(* IEC 61131-3 sources: PO_LAB_3/Physical/Acp10_MC (part 2) *)

(* ---- acp10_mc.fun ---- *)
FUNCTION_BLOCK MC_AbortTrigger (*aborts FBs connected to trigger events*)
	VAR_INPUT
		Axis : UDINT; (*axis reference, defines on which axis the trigger should be aborted*)
		TriggerInput : MC_TRIGGER_REF; (*trigger input signal source*)
		Execute : BOOL; (*aborts the trigger at rising edge*)
	END_VAR
	VAR_OUTPUT
		Done : BOOL; (*FB with trigger has been aborted*)
		Busy : BOOL; (*the function block is not finished*)
		Error : BOOL; (*error occurred in FB*)
		ErrorID : UINT; (*error number*)
	END_VAR
	VAR
		C_Axis : UDINT; (*internal variable*)
		state : USINT; (*internal variable*)
		C_Done : BOOL; (*internal variable*)
		C_Error : BOOL; (*internal variable*)
		C_ErrorID : UINT; (*internal variable*)
	END_VAR
END_FUNCTION_BLOCK

FUNCTION_BLOCK MC_BR_AutCommand (*transferes commands for the cam automat to the drive*)
	VAR_INPUT
		Slave : UDINT; (*axis reference of the slave axis*)
		Enable : BOOL; (*activates the function block*)
		Start : BOOL; (*starts the cam automat*)
		Stop : BOOL; (*stops the movement on the slave axis*)
		Deceleration : REAL; (*deceleration for the stop command*)
		Restart : BOOL; (*reengages the slave axis to the automat*)
		EndAutomat : BOOL; (*aborts the automat in the background*)
		SetSignal1 : BOOL; (*sets the automat signal1*)
		SetSignal2 : BOOL; (*sets the automat signal2*)
		SetSignal3 : BOOL; (*sets the automat signal3*)
		SetSignal4 : BOOL; (*sets the automat signal4*)
		ResetSignal1 : BOOL; (*resets the automat signal1*)
		ResetSignal2 : BOOL; (*resets the automat signal2*)
		ResetSignal3 : BOOL; (*resets the automat signal3*)
		ResetSignal4 : BOOL; (*resets the automat signal4*)
		TransferParLock : BOOL; (*transfer the par lock parameter*)
		SelectParLock : USINT; (*select the par lock parameter*)
	END_VAR
	VAR_OUTPUT
		Active : BOOL; (*function block is active and waits for command*)
		Busy : BOOL; (*function block is enabled*)
		CommandAborted : BOOL; (*function block was aborted by another function block*)
		Error : BOOL; (*error occurred in the function block*)
		ErrorID : UINT; (*error number*)
		Running : BOOL; (*slave is engaged to the automat*)
		StandBy : BOOL; (*cam automat is active in the background*)
		ParLockTransferred : BOOL; (*par lock parameter transferred*)
		ActualStateIndex : USINT; (*actual state of the cam automat*)
		ActualStateCamIndex : UINT; (*actual cam index of the actual state*)
		InCam : BOOL; (*automat is in cam*)
		InCompensation : BOOL; (*automat is in compensation*)
	END_VAR
	VAR
		C_Slave : UDINT; (*internal variable*)
		IS : MC_0099_IS_TYP; (*internal variable*)
	END_VAR
END_FUNCTION_BLOCK

FUNCTION_BLOCK MC_BR_AutControl (*controls the cam automat functions*)
	VAR_INPUT
		Enable : BOOL; (*enables the functionality of this FB*)
		Slave : UDINT; (*axis reference of the slave axis*)
		ParLock : USINT; (*lock for consistent online change*)
		Signal1 : BOOL; (*set signal1*)
		Signal2 : BOOL; (*set signal2*)
		Signal3 : BOOL; (*set signal3*)
		Signal4 : BOOL; (*set signal4*)
		Start : BOOL; (*start automat*)
		Stop : BOOL; (*stop automat*)
		Deceleration : REAL; (*deceleration for stop command*)
		Restart : BOOL; (*restart command*)
		AdrAutData : UDINT; (*address of optional cam automat data structure*)
		InitAutData : BOOL; (*initialize the parameters of the optional cam automat data structure*)
	END_VAR
	VAR_OUTPUT
		Active : BOOL; (*automat control function block activated*)
		Busy : BOOL; (*function block is not finished*)
		Error : BOOL; (*error occurred in FB*)
		ErrorID : UINT; (*error number*)
		AutDataInitialized : BOOL; (*cam automat data structure initialized*)
		Running : BOOL; (*cam automat is running*)
		ActualStateIndex : USINT; (*index of the actual state*)
		ActualCamType : USINT; (*cam type of the actual state*)
	END_VAR
	VAR
		C_Slave : UDINT; (*internal variable*)
		ParLockOld : USINT; (*internal variable*)
		LockID : USINT; (*internal variable*)
		CmdParLock : BOOL; (*internal variable*)
		EdgeSignal1 : BOOL; (*internal variable*)
		EdgeSignal2 : BOOL; (*internal variable*)
		EdgeSignal3 : BOOL; (*internal variable*)
		EdgeSignal4 : BOOL; (*internal variable*)
		EdgeStart : BOOL; (*internal variable*)
		CmdStart : BOOL; (*internal variable*)
		EdgeStop : BOOL; (*internal variable*)
		CmdStop : BOOL; (*internal variable*)
		C_Deceleration : REAL; (*internal variable*)
		EdgeRestart : BOOL; (*internal variable*)
		CmdRestart : BOOL; (*internal variable*)
		EdgeInitAutData : BOOL; (*internal variable*)
		CmdInitAutData : BOOL; (*internal variable*)
		C_AutData : MC_AUTDATA_TYP; (*internal variable*)
		C_Master : UDINT; (*internal variable*)
		C_Error : BOOL; (*internal variable*)
		C_ErrorID : UINT; (*internal variable*)
		CC_ErrorID : UINT; (*internal variable*)
		SignalSet : USINT; (*internal variable*)
		SignalReset : USINT; (*internal variable*)
		CmdAutStart : UINT; (*internal variable*)
		AutStatusValid : BOOL; (*internal variable*)
		AutStateDld : USINT; (*internal variable*)
		AutStatusOffset : UINT; (*internal variable*)
		AutStatusRecIndex : USINT; (*internal variable*)
		LockIDSend : USINT; (*internal variable*)
		AutActualStateIndexOffset : UINT; (*internal variable*)
		AutActualStateIndexRecIndex : USINT; (*internal variable*)
		C_Busy : BOOL; (*internal variable*)
		AutActualCamTypeOffset : UINT; (*internal variable*)
		AutActualCamTypeRecIndex : USINT; (*internal variable*)
		LockIDMa : USINT; (*internal variable*)
		sendSlot : USINT; (*internal variable*)
		readSlot : USINT; (*internal variable*)
		state : USINT; (*internal variable*)
		LockIDPar : USINT; (*internal variable*)
		MoveID : USINT; (*internal variable*)
		LockIDReceive : USINT; (*internal variable*)
	END_VAR
END_FUNCTION_BLOCK

FUNCTION_BLOCK MC_BR_AutoCamDwell (*starts a link between master and slave with a self calculated cam profile*)
	VAR_INPUT
		Master : UDINT; (*axis reference of the master axis*)
		Slave : UDINT; (*axis reference of the slave axis*)
		Enable : BOOL; (*function block is activated*)
		InitData : BOOL; (*start transferring the parameters*)
		LeadInMasterDistance : REAL; (*master axis compensation distance for the lead in*)
		LeadInSlaveDistance : REAL; (*slave axis compensation distance for the lead in*)
		LeadOutMasterDistance : REAL; (*master axis compensation distance for the lead out*)
		LeadOutSlaveDistance : REAL; (*slave axis compensation distance for the lead out*)
		MasterStartPosition : REAL; (*master position where the cam profile starts*)
		MasterDwellDistance : REAL; (*master length of the optional dwell section*)
		MasterLength : REAL; (*master side length of the automatically calculated cam profile*)
		SlaveLength : REAL; (*slave side length of the automatically calculated cam profile*)
		MasterParID : UINT; (*use this ParID for the master axis instead of the set position*)
		MasterParIDMaxVelocity : REAL; (*maximum speed of the master ParID value*)
		LeadInSignal : BOOL; (*signal from the control to start the lead in*)
		LeadOutSignal : BOOL; (*signal from the control to start the lead out*)
		LeadInParID : UINT; (*ParID that can be used by the drive to start the lead in*)
		LeadOutParID : UINT; (*ParID that can be used by the drive to start the lead out*)
	END_VAR
	VAR_OUTPUT
		Active : BOOL; (*parameters are transferred and FB is active*)
		Busy : BOOL; (*function block is enabled*)
		CommandAborted : BOOL; (*function block aborted by another FB*)
		Error : BOOL; (*error occurred in FB*)
		ErrorID : UINT; (*error number*)
		DataInitialized : BOOL; (*parameters are transferred*)
		InSync : BOOL; (*cam profile is synchronized with the master*)
		InCam : BOOL; (*the coupling is within the cam range*)
		InDwell : BOOL; (*the coupling is within the dwell range*)
	END_VAR
	VAR
		C_Master : UDINT; (*internal variable*)
		C_Slave : UDINT; (*internal variable*)
		EdgeInitData : BOOL; (*internal variable*)
		C_LeadInMasterDistance : DINT; (*internal variable*)
		C_LeadInSlaveDistance : DINT; (*internal variable*)
		C_LeadOutMasterDistance : DINT; (*internal variable*)
		C_LeadOutSlaveDistance : DINT; (*internal variable*)
		C_MasterStartPosition : DINT; (*internal variable*)
		C_MasterDwellDistance : DINT; (*internal variable*)
		C_MasterLength : DINT; (*internal variable*)
		C_SlaveLength : DINT; (*internal variable*)
		C_MasterParID : UINT; (*internal variable*)
		C_MasterParIDMaxVelocity : REAL; (*internal variable*)
		C_LeadInParID : UINT; (*internal variable*)
		C_LeadOutParID : UINT; (*internal variable*)
		EdgeLeadInSignal : BOOL; (*internal variable*)
		EdgeLeadOutSignal : BOOL; (*internal variable*)
		LeadInSignalUsed : BOOL; (*internal variable*)
		LeadOutSignalUsed : BOOL; (*internal variable*)
		C_Active : BOOL; (*internal variable*)
		C_Busy : BOOL; (*internal variable*)
		C_CommandAborted : BOOL; (*internal variable*)
		C_Error : BOOL; (*internal variable*)
		C_ErrorID : UINT; (*internal variable*)
		CC_ErrorID : UINT; (*internal variable*)
		C_InSync : BOOL; (*internal variable*)
		C_InCam : BOOL; (*internal variable*)
		C_InDwell : BOOL; (*internal variable*)
		RunningMasterDwellDistance : DINT; (*internal variable*)
		ArithIndex : UINT; (*internal variable*)
		CmpIndex : UINT; (*internal variable*)
		MuxIndex : UINT; (*internal variable*)
		EvWrIndex : UINT; (*internal variable*)
		VarIndex : UINT; (*internal variable*)
		LogicIndex : UINT; (*internal variable*)
		AutStatusValid : BOOL; (*internal variable*)
		AutActualStateIndexOffset : UINT; (*internal variable*)
		AutActualStateIndexRecIndex : USINT; (*internal variable*)
		LockIDMa : USINT; (*internal variable*)
		sendSlot : USINT; (*internal variable*)
		readSlot : USINT; (*internal variable*)
		state : USINT; (*internal variable*)
		LockID : USINT; (*internal variable*)
		LockIDPar : USINT; (*internal variable*)
		LockIDSend : USINT; (*internal variable*)
		MoveID : USINT; (*internal variable*)
		LockIDReceive : USINT; (*internal variable*)
	END_VAR
END_FUNCTION_BLOCK

FUNCTION_BLOCK MC_BR_AxisErrorCollector (*collects information if a FB or axis error occured and if an axis is in state Errorstop*)
	VAR_INPUT
		Axis : UDINT; (*axis reference*)
		Enable : BOOL; (*function block is activated*)
	END_VAR
	VAR_OUTPUT
		Valid : BOOL; (*if set, the data of the other outputs is valid*)
		Busy : BOOL; (*function block is not finished*)
		Error : BOOL; (*error occurred in FB*)
		ErrorID : UINT; (*error number*)
		FunctionBlockError : BOOL; (*at least one function block reported an error*)
		AxisError : BOOL; (*at least one axis error was reported*)
		AxisWarning : BOOL; (*at least one axis warning was reported*)
		Errorstop : BOOL; (*the axis is in state Errorstop*)
	END_VAR
	VAR
		C_Axis : UDINT; (*internal variable*)
		IS : MC_0104_IS_TYP; (*internal variable*)
	END_VAR
END_FUNCTION_BLOCK

FUNCTION_BLOCK MC_BR_BrakeControl (*executes several commands for holding brake*)
	VAR_INPUT
		Axis : UDINT; (*axis reference*)
		Execute : BOOL; (*execute brake command at rising edge*)
		Command : USINT; (*brake command*)
		Configuration : MC_BRAKE_CONFIG_REF; (*brake configuration*)
	END_VAR
	VAR_OUTPUT
		Done : BOOL; (*brake command done*)
		Busy : BOOL; (*function block is not finished*)
		Error : BOOL; (*error occured in FB*)
		ErrorID : UINT; (*error number*)
		PositionError : REAL; (*position error of holding brake test*)
		BrakeStatus : BOOL; (*actual brake status*)
	END_VAR
	VAR
		C_Axis : UDINT; (*internal variable*)
		IS : MC_0110_IS_TYP; (*internal variable*)
	END_VAR
END_FUNCTION_BLOCK

FUNCTION_BLOCK MC_BR_BrakeOperation (*opens and closes the holding brake when the controller is off*)
	VAR_INPUT
		Axis : UDINT; (*axis reference*)
		Execute : BOOL; (*execute brake command at rising edge*)
		BrakeCommand : USINT; (*brake command, open or close*)
	END_VAR
	VAR_OUTPUT
		Done : BOOL; (*brake command done*)
		Busy : BOOL; (*function block is not finished*)
		Error : BOOL; (*error occurred in FB*)
		ErrorID : UINT; (*error number*)
	END_VAR
	VAR
		C_Axis : UDINT; (*internal variable*)
		C_Execute : BOOL; (*internal variable*)
		C_BrakeCommand : USINT; (*internal variable*)
		C_Done : BOOL; (*internal variable*)
		LockIDPar : USINT; (*internal variable*)
		C_ErrorID : UINT; (*internal variable*)
		C_Error : BOOL; (*internal variable*)
		state : USINT; (*internal variable*)
	END_VAR
END_FUNCTION_BLOCK

FUNCTION_BLOCK MC_BR_CalcCamFromPoints (*calculates a cam profile from a list of points*)
	VAR_INPUT
		Execute : BOOL; (*calculation starts at rising edge*)
		MasterPointsAddress : UDINT; (*data address of the master points list*)
		SlavePointsAddress : UDINT; (*data address of the slave points list*)
		NumberOfPoints : UINT; (*number of master and slave points*)
		CamProfileAddress : UDINT; (*data address for the calculated cam profile*)
		Configuration : MC_CALC_CAM_CONFIG_REF; (*optional additional configuration*)
	END_VAR
	VAR_OUTPUT
		Done : BOOL; (*calculation is complete*)
		Busy : BOOL; (*function block is not finished*)
		Error : BOOL; (*error occurred in FB*)
		ErrorID : UINT; (*error number*)
	END_VAR
	VAR
		IS : MC_0093_IS_TYP; (*internal variable*)
	END_VAR
END_FUNCTION_BLOCK

FUNCTION_BLOCK MC_BR_CalcCamFromSections (*calculates from a list of points a cam profile*)
	VAR_INPUT
		Execute : BOOL; (*calculation starts at rising edge*)
		DataAddress : UDINT; (*data address of the input data with the list of points*)
		CamProfileAddress : UDINT; (*data address for the calculated cam profile*)
	END_VAR
	VAR_OUTPUT
		Done : BOOL; (*calculation is complete*)
		Busy : BOOL; (*function block is not finished*)
		Error : BOOL; (*error occurred in FB*)
		ErrorID : UINT; (*error number*)
		ErrorInSection : UINT; (*index of section with error*)
	END_VAR
	VAR
		C_ErrorID : UINT; (*internal variable*)
		C_ErrorInSection : UINT; (*internal variable*)
		C_Error : BOOL; (*internal variable*)
		state : USINT; (*internal variable*)
	END_VAR
END_FUNCTION_BLOCK

FUNCTION_BLOCK MC_BR_CalcPointsFromCam (*calculates a list of points from a cam profile*)
	VAR_INPUT
		Execute : BOOL; (*calculation starts at rising edge*)
		DataObjectName : STRING[12]; (*name of the cam table*)
		MasterPointsAddress : UDINT; (*data address of the master points list*)
		SlavePointsAddress : UDINT; (*data address of the slave points list*)
		NumberOfPoints : UINT; (*number of master and slave points*)
	END_VAR
	VAR_OUTPUT
		Done : BOOL; (*calculation is complete*)
		Busy : BOOL; (*function block is not finished *)
		Error : BOOL; (*error occured in FB*)
		ErrorID : UINT; (*error number*)
		AdditionalInfo : MC_CALC_CAM_CONFIG_REF; (*additional information about the cam profile*)
	END_VAR
	VAR
		IS : MC_0123_IS_TYP; (*internal variable*)
	END_VAR
END_FUNCTION_BLOCK

FUNCTION_BLOCK MC_BR_CalcSectionsFromCam (*calculates the sections from a cam profile *)
	VAR_INPUT
		Execute : BOOL; (*calculation starts at rising edge*)
		DataObjectName : STRING[12]; (*name of the cam table*)
		DataAddress : UDINT; (*address of the variable for the sections*)
	END_VAR
	VAR_OUTPUT
		Done : BOOL; (*calculation is complete*)
		Busy : BOOL; (*function block is not finished *)
		Error : BOOL; (*error occured in FB*)
		ErrorID : UINT; (*error number*)
	END_VAR
	VAR
		IS : MC_0122_IS_TYP; (*internal variable*)
	END_VAR
END_FUNCTION_BLOCK

FUNCTION_BLOCK MC_BR_CamIn (*starts a cam profile link between the master and the slave axis*)
	VAR_INPUT
		Master : UDINT; (*axis reference of the master axis*)
		Slave : UDINT; (*axis reference of the slave axis*)
		Enable : BOOL; (*function block is activated*)
		InitData : BOOL; (*starts transferring the parameters*)
		CamTableID : USINT; (*ID number of the cam profile*)
		MasterStartPosition : REAL; (*master position where the cam profile starts*)
		MasterScaling : DINT; (*factor of the master profile*)
		SlaveScaling : DINT; (*factor of the slave scaling*)
		EnterCam : BOOL; (*signal from the control to start the coupling*)
		ExitCam : BOOL; (*signal from the control to end the coupling*)
		Restart : BOOL; (*signal from the control to restart the coupling*)
        AdvancedParameters: MC_ADVANCED_CAM_PAR_REF; (*additional inputs for advanced usage of FB*)
	END_VAR
	VAR_OUTPUT
		Active : BOOL; (*parameters are transferred and FB is active*)
		Busy : BOOL; (*function block is enabled*)
		CommandAborted : BOOL; (*function block aborted by another FB*)
		Error : BOOL; (*error occurred in FB*)
		ErrorID : UINT; (*error number*)
		DataInitialized : BOOL; (*transferring parameters is completed*)
		Running : BOOL; (*cam coupling is running*)
		StandBy : BOOL; (*cam coupling is active in the background*)
		InLeadIn : BOOL; (*the coupling is within the leadin range*)
		InCam : BOOL; (*the coupling is within the cam range*)
		InLeadOut : BOOL; (*the coupling is within the leadout range*)
		EndOfProfile : BOOL; (*pulsed output signaling the cyclic end of the cam profile*)
	END_VAR
	VAR
		C_Master : UDINT; (*internal variable*)
		C_Slave : UDINT; (*internal variable*)
		IS: MC_0146_IS_TYP; (*internal variable*)
	END_VAR
END_FUNCTION_BLOCK

FUNCTION_BLOCK MC_BR_CamDwell (*starts a cam profile link between the master and the slave axis*)
	VAR_INPUT
		Master : UDINT; (*axis reference of the master axis*)
		Slave : UDINT; (*axis reference of the slave axis*)
		Enable : BOOL; (*function block is activated*)
		InitData : BOOL; (*starts transferring the parameters*)
		LeadInMasterDistance : REAL; (*master axis compensation distance for the lead in*)
		LeadInSlaveDistance : REAL; (*slave axis compensation distance for the lead in*)
		LeadInMasterOffset : REAL; (*master side offset within the cam profile*)
		LeadOutMasterDistance : REAL; (*master axis compensation distance for the lead out*)
		LeadOutSlaveDistance : REAL; (*slave axis compensation distance for the lead out*)
		LeadOutMasterOffset : REAL; (*master side offset within the cam profile*)
		MasterStartPosition : REAL; (*master position where the cam profile starts*)
		MasterDwellDistance : REAL; (*master length of the optional dwell section*)
		MasterScaling : REAL; (*factor of the master profile*)
		SlaveScaling : REAL; (*factor of the slave scaling*)
		CamTableID : USINT; (*ID number of the cam profile*)
		MasterParID : UINT; (*use this ParID for the master axis instead of the set position*)
		MasterParIDMaxVelocity : REAL; (*maximum speed of the master ParID value*)
		LeadInSignal : BOOL; (*signal from the control to start the lead in*)
		LeadOutSignal : BOOL; (*signal from the control to start the lead out*)
		LeadInParID : UINT; (*ParID that can be used by the drive to start the lead out movement*)
		LeadOutParID : UINT; (*ParID that can be used by the drive to start the lead out movement*)
	END_VAR
	VAR_OUTPUT
		Active : BOOL; (*parameters are transferred and FB is active*)
		Busy : BOOL; (*function block is enabled*)
		CommandAborted : BOOL; (*function block aborted by another FB*)
		Error : BOOL; (*error occurred in FB*)
		ErrorID : UINT; (*error number*)
		DataInitialized : BOOL; (*transferring parameters is completed*)
		InSync : BOOL; (*cam profile is synchronized with the master*)
		InCam : BOOL; (*the coupling is within the cam range*)
		InDwell : BOOL; (*the coupling is within the dwell range*)
	END_VAR
	VAR
		C_Master : UDINT; (*internal variable*)
		C_Slave : UDINT; (*internal variable*)
		EdgeInitData : BOOL; (*internal variable*)
		C_LeadInMasterDistance : DINT; (*internal variable*)
		C_LeadInSlaveDistance : DINT; (*internal variable*)
		C_LeadInMasterOffset : DINT; (*internal variable*)
		C_LeadOutMasterDistance : DINT; (*internal variable*)
		C_LeadOutSlaveDistance : DINT; (*internal variable*)
		C_LeadOutMasterOffset : DINT; (*internal variable*)
		C_MasterStartPosition : DINT; (*internal variable*)
		C_MasterDwellDistance : DINT; (*internal variable*)
		C_MasterScaling : DINT; (*internal variable*)
		C_SlaveScaling : DINT; (*internal variable*)
		C_CamTableID : UINT; (*internal variable*)
		C_MasterParID : UINT; (*internal variable*)
		C_MasterParIDMaxVelocity : REAL; (*internal variable*)
		C_LeadInParID : UINT; (*internal variable*)
		C_LeadOutParID : UINT; (*internal variable*)
		EdgeLeadInSignal : BOOL; (*internal variable*)
		EdgeLeadOutSignal : BOOL; (*internal variable*)
		LeadInSignalUsed : BOOL; (*internal variable*)
		LeadOutSignalUsed : BOOL; (*internal variable*)
		C_Active : BOOL; (*internal variable*)
		C_Busy : BOOL; (*internal variable*)
		C_CommandAborted : BOOL; (*internal variable*)
		C_Error : BOOL; (*internal variable*)
		C_ErrorID : UINT; (*internal variable*)
		CC_ErrorID : UINT; (*internal variable*)
		C_InSync : BOOL; (*internal variable*)
		C_InCam : BOOL; (*internal variable*)
		C_InDwell : BOOL; (*internal variable*)
		RunningMasterDwellDistance : DINT; (*internal variable*)
		ArithIndex : UINT; (*internal variable*)
		CmpIndex : UINT; (*internal variable*)
		MuxIndex : UINT; (*internal variable*)
		EvWrIndex : UINT; (*internal variable*)
		VarIndex : UINT; (*internal variable*)
		LogicIndex : UINT; (*internal variable*)
		AutStatusValid : BOOL; (*internal variable*)
		AutActualStateIndexOffset : UINT; (*internal variable*)
		AutActualStateIndexRecIndex : USINT; (*internal variable*)
		LockIDMa : USINT; (*internal variable*)
		AutActualCamTypeOffset : UINT; (*internal variable*)
		AutActualCamTypeRecIndex : USINT; (*internal variable*)
		LockIDSend : USINT; (*internal variable*)
		sendSlot : USINT; (*internal variable*)
		readSlot : USINT; (*internal variable*)
		state : USINT; (*internal variable*)
		LockID : USINT; (*internal variable*)
		LockIDPar : USINT; (*internal variable*)
		LockIDReceive : USINT; (*internal variable*)
		MoveID : USINT; (*internal variable*)
	END_VAR
END_FUNCTION_BLOCK

FUNCTION_BLOCK MC_BR_CamTransition (*starts a cam profile link between the master and the slave axis*)
	VAR_INPUT
		Master : UDINT; (*axis reference of the master axis*)
		Slave : UDINT; (*axis reference of the slave axis*)
		Enable : BOOL; (*function block is activated*)
		InitData : BOOL; (*starts transferring the parameters*)
		LeadInMasterDistance : REAL; (*master axis compensation distance for the lead in*)
		LeadInSlaveDistance : REAL; (*slave axis compensation distance for the lead in*)
		LeadInMasterOffset : REAL; (*master side offset within the cam profile*)
		LeadOutMasterDistance : REAL; (*master axis compensation distance for the lead out*)
		LeadOutSlaveDistance : REAL; (*slave axis compensation distance for the lead out*)
		LeadOutMasterOffset : REAL; (*master side offset within the cam profile*)
		ReverseSlaveDistance : REAL; (*slaves moves this distence in reverse direction during transition*)
		MasterInterval : REAL; (*interval length of master movement: cam + transition*)
		SlaveInterval : REAL; (*interval length of slave movement: cam + transition*)
		MasterStartPosition : REAL; (*master position where the cam profile starts*)
		MasterScaling : REAL; (*factor of the master profile*)
		SlaveScaling : REAL; (*factor of the slave scaling*)
		CamTableID : USINT; (*ID number of the cam profile*)
		MasterParID : UINT; (*use this ParID for the master axis instead of the set position*)
		MasterParIDMaxVelocity : REAL; (*maximum speed of the master ParID value*)
		LeadInSignal : BOOL; (*signal from the control to start the lead in*)
		LeadOutSignal : BOOL; (*signal from the control to start the lead out*)
		LeadInParID : UINT; (*ParID that can be used by the drive to start the lead out movement*)
		LeadOutParID : UINT; (*ParID that can be used by the drive to start the lead out movement*)
		TransitionMode : UINT; (*mode for transition movement*)
		CamMode : UINT; (*mode for cam movement*)
		CamTime : REAL; (*time for cam movement in mode mcTIME_BASED*)
	END_VAR
	VAR_OUTPUT
		Active : BOOL; (*parameters are transferred and FB is active*)
		Busy : BOOL; (*function block is enabled*)
		CommandAborted : BOOL; (*function block aborted by another FB*)
		Error : BOOL; (*error occurred in FB*)
		ErrorID : UINT; (*error number*)
		DataInitialized : BOOL; (*transferring parameters is completed*)
		InSync : BOOL; (*cam profile is synchronized with the master*)
		InLeadIn : BOOL; (*the coupling is within the leadin range*)
		InCam : BOOL; (*the coupling is within the cam range*)
		InTransition : BOOL; (*the coupling is within the transition range*)
		InReverse : BOOL; (*the coupling is within the reverse reange*)
		InLeadOut : BOOL; (*the coupling is within the leadout range*)
	END_VAR
	VAR
		C_Master : UDINT; (*internal variable*)
		C_Slave : UDINT; (*internal variable*)
		EdgeInitData : BOOL; (*internal variable*)
		C_LeadInMasterDistance : DINT; (*internal variable*)
		C_LeadInSlaveDistance : DINT; (*internal variable*)
		C_LeadInMasterOffset : DINT; (*internal variable*)
		C_LeadOutMasterDistance : DINT; (*internal variable*)
		C_LeadOutSlaveDistance : DINT; (*internal variable*)
		C_LeadOutMasterOffset : DINT; (*internal variable*)
		C_ReverseSlaveDistance : DINT; (*internal variable*)
		C_MasterInterval : DINT; (*internal variable*)
		C_SlaveInterval : DINT; (*internal variable*)
		C_MasterStartPosition : DINT; (*internal variable*)
		C_MasterScaling : DINT; (*internal variable*)
		C_SlaveScaling : DINT; (*internal variable*)
		C_CamTableID : UINT; (*internal variable*)
		C_MasterParID : UINT; (*internal variable*)
		C_MasterParIDMaxVelocity : REAL; (*internal variable*)
		C_LeadInParID : UINT; (*internal variable*)
		C_LeadOutParID : UINT; (*internal variable*)
		C_TransitionMode : UINT; (*internal variable*)
		C_CamMode : UINT; (*internal variable*)
		C_CamTime : REAL; (*internal variable*)
		EdgeLeadInSignal : BOOL; (*internal variable*)
		EdgeLeadOutSignal : BOOL; (*internal variable*)
		LeadInSignalUsed : BOOL; (*internal variable*)
		LeadOutSignalUsed : BOOL; (*internal variable*)
		C_Active : BOOL; (*internal variable*)
		C_Busy : BOOL; (*internal variable*)
		C_CommandAborted : BOOL; (*internal variable*)
		C_Error : BOOL; (*internal variable*)
		C_ErrorID : UINT; (*internal variable*)
		CC_ErrorID : UINT; (*internal variable*)
		C_InSync : BOOL; (*internal variable*)
		C_InCam : BOOL; (*internal variable*)
		C_InTransition : BOOL; (*internal variable*)
		C_InReverse : BOOL; (*internal variable*)
		C_InLeadIn : BOOL; (*internal variable*)
		C_InLeadOut : BOOL; (*internal variable*)
		C_MasterCompDistance : DINT; (*internal variable*)
		C_SlaveCompDistance : DINT; (*internal variable*)
		C_OldMasterCompDistance : DINT; (*internal variable*)
		C_OldSlaveCompDistance : DINT; (*internal variable*)
		C_CamMasterPeriod : DINT; (*internal variable*)
		C_CamSlavePeriod : DINT; (*internal variable*)
		ArithIndex : UINT; (*internal variable*)
		CmpIndex : UINT; (*internal variable*)
		MuxIndex : UINT; (*internal variable*)
		EvWrIndex : UINT; (*internal variable*)
		VarIndex : UINT; (*internal variable*)
		LogicIndex : UINT; (*internal variable*)
		PidIndex : UINT; (*internal variable*)
		AutStatusValid : BOOL; (*internal variable*)
		InitDataUsed : BOOL; (*internal variable*)
		AutActualStateIndexOffset : UINT; (*internal variable*)
		AutActualStateIndexRecIndex : USINT; (*internal variable*)
		oldAutomatState : USINT; (*internal variable*)
		MasterVelocityOffset : UINT; (*internal variable*)
		MasterVelocityRecIndex : USINT; (*internal variable*)
		LockIDMa : USINT; (*internal variable*)
		AutActualCamTypeOffset : UINT; (*internal variable*)
		AutActualCamTypeRecIndex : USINT; (*internal variable*)
		ChangePending : BOOL; (*internal variable*)
		sendSlot : USINT; (*internal variable*)
		readSlot : USINT; (*internal variable*)
		state : USINT; (*internal variable*)
		LockID : USINT; (*internal variable*)
		LockIDPar : USINT; (*internal variable*)
		MoveID : USINT; (*internal variable*)
		LockIDSend : USINT; (*internal variable*)
		Reserve3 : UDINT; (*internal variable*)
		nextState : USINT; (*internal variable*)
		Reserve4 : USINT; (*internal variable*)
		LockIDReceive : USINT; (*internal variable*)
		Reserve6 : BOOL; (*internal variable*)
	END_VAR
END_FUNCTION_BLOCK

FUNCTION_BLOCK MC_BR_CheckAutCompensation (*checks the compensation data of a cam profile automat*)
	VAR_INPUT
		Master : UDINT; (*axis reference of the master axis*)
		Slave : UDINT; (*axis reference of the slave axis*)
		Execute : BOOL; (*check the compensation data at rising edge*)
		Mode : UINT; (*choose the mode*)
		CompensationData : MC_AUT_COMP_DATA_REF; (*compensation data for the check or calculation*)
	END_VAR
	VAR_OUTPUT
		Done : BOOL; (*check or calculation is successfully finished*)
		Busy : BOOL; (*function block is not finished yet*)
		Error : BOOL; (*error occured in FB*)
		ErrorID : UINT; (*error number*)
		Result : REAL; (*result of the calculation*)
	END_VAR
	VAR
		C_Master : UDINT; (*internal variable*)
		C_Slave : UDINT; (*internal variable*)
		IS : MC_0103_IS_TYP; (*internal variable*)
	END_VAR
END_FUNCTION_BLOCK

FUNCTION_BLOCK MC_BR_CheckEndlessPosition (*checks the endless position data for restoring the axis position*)
	VAR_INPUT
		Axis : UDINT; (*axis reference*)
		Execute : BOOL; (*check the endless position data at rising edge*)
		DataAddress : UDINT; (*data address of momory storage for endless position*)
	END_VAR
	VAR_OUTPUT
		Done : BOOL; (*memory storage for endless position was checked*)
		Busy : BOOL; (*function block is not finished*)
		Error : BOOL; (*error occurred in FB*)
		ErrorID : UINT; (*error number*)
		EndlessPositionInitialized : BOOL; (*address of memory storage already initialized*)
		DataValid : BOOL; (*axis position can be restored from the endless position data*)
	END_VAR
	VAR
		C_Axis : UDINT; (*internal variable*)
		IS : MC_0130_IS_TYP; (*internal variable*)
	END_VAR
END_FUNCTION_BLOCK

FUNCTION_BLOCK MC_BR_CommandError (*transfers error commands to the drive, where they are entered*)
	VAR_INPUT
		Axis  : UDINT; (*axis reference*)
		Execute : BOOL; (*transfer command at rising edge*)
		Command : UINT; (*error command*)
	END_VAR
	VAR_OUTPUT
		Done  : BOOL; (*command was successfully transferred *)
		Busy  : BOOL; (*function block is not finished yet*)
		Error : BOOL; (*error occured in FB*)
		ErrorID : UINT; (*error number *)
	END_VAR
	VAR
		C_Axis : UDINT; (*internal variable*)
		IS : MC_0140_IS_TYP; (*internal variable*)
	END_VAR
END_FUNCTION_BLOCK

FUNCTION_BLOCK MC_BR_ConfigPowerStageCheck (*configurates the power stage checks of the ACOPOS*)
	VAR_INPUT
		Axis : UDINT; (*axis reference*)
		Execute : BOOL; (*transfer configuration at rising edge *)
		Configuration : MC_POWER_STAGE_CHECK_REF; (*configuration data*)
	END_VAR
	VAR_OUTPUT
		Done : BOOL; (*configuration is successfully finished*)
		Busy : BOOL; (*function block is not finished yet*)
		Error : BOOL; (*error occured in FB*)
		ErrorID : UINT; (*error number*)
	END_VAR
	VAR
		C_Axis : UDINT; (*internal variable*)
		IS : MC_0137_IS_TYP; (*internal variable*)
	END_VAR
END_FUNCTION_BLOCK

FUNCTION_BLOCK MC_BR_CrossCutterControl (*controls a cutter axis linked to a master axis*)
	VAR_INPUT
		Master : UDINT; (*axis reference of the master axis*)
		Slave : UDINT; (*axis reference of the slave/cutter axis*)
		Enable : BOOL; (*function block is activated*)
		InitData : BOOL; (*starts transferring the parameters*)
		EnableCut : BOOL; (*start/stop synchronizing slave to master*)
		CutRangeMaster : REAL; (*cut area on master axis, where the cutter needs to run synchronous to master*)
		CutRangeSlave : REAL; (*area around cut point on slave axis, where the cutter needs to run synchronous to master*)
		ProductLength : REAL; (*distance (master based) in which the cutter needs to make one cut*)
		ProductLengthCorrection : REAL; (*this value is added to ProductLength and then downloaded*)
		AdvancedParameters : MC_ADVANCED_CUT_PAR_REF; (*additional inputs for advanced usage of FB*)
	END_VAR
	VAR_OUTPUT
		Active : BOOL; (*parameters are transferred and FB is active*)
		Busy : BOOL; (*function block is enabled*)
		CommandAborted : BOOL; (*function block aborted by another FB*)
		Error : BOOL; (*error occurred in FB*)
		ErrorID : UINT; (*error number*)
		DataInitialized : BOOL; (*transferring parameters is completed*)
		StandBy : BOOL; (*FB can be restarted*)
		InCompensation : BOOL; (*axis outside CutRange, and synchronized*)
		InCut : BOOL; (*axis is within CutRange*)
		CutCount : UDINT; (*information about how many cuts have been made*)
		CutMasterPosition : DINT; (*latched master position at cut for registration mark control*)
	END_VAR
	VAR
		C_Master : UDINT; (*internal variable*)
		C_Slave : UDINT; (*internal variable*)
		IS : MC_0114_IS_TYP; (*internal variable*)
	END_VAR
END_FUNCTION_BLOCK

FUNCTION_BLOCK MC_BR_CyclicRead (*enters the specified ParID in the cyclic data from drive and returns it*)
	VAR_INPUT
		Axis : UDINT; (*axis reference*)
		Enable : BOOL; (*specified ParID is read from the drive as long as enable is TRUE*)
		ParID : UINT; (*ParID which should be read from the drive*)
		DataAddress : UDINT; (*data address of the variable for the value of the ParID*)
		DataType : UINT; (*data type of the ParID*)
		Mode : UINT; (*mode for configuration of records*)
	END_VAR
	VAR_OUTPUT
		Valid : BOOL; (*when set the output is valid*)
		Busy : BOOL; (*function block is not finished*)
		Error : BOOL; (*error occurred in FB*)
		ErrorID : UINT; (*error number*)
	END_VAR
	VAR
		C_Axis : UDINT; (*internal variable*)
		IS : MC_0069_IS_TYP; (*internal variable*)
	END_VAR
END_FUNCTION_BLOCK

FUNCTION_BLOCK MC_BR_CyclicReadDataInfo (*Read administrative information of cyclic read data*)
	VAR_INPUT
		Axis : UDINT; (*axis reference*)
		Enable : BOOL; (*function block is activated*)
	END_VAR
	VAR_OUTPUT
		Valid : BOOL; (*if set, the data of the other outputs is valid*)
		Busy : BOOL; (*function block is not finished*)
		Error : BOOL; (*error occurred in FB*)
		ErrorID : UINT; (*error number*)
		RecordCount : UINT; (*number of configured records from the drive*)
		ParIDCount : UINT; (*number of configured ParIDs from the drive*)
		RecordUpdateTime : DINT; (*update time of one single record from the drive*)
		TotalUpdateTime : DINT; (*update time of all records from the drive*)
		RecordIndex : UINT; (*index of currently read record from the drive*)
		RecordInfo : MC_RECORD_INFO_REF; (*detailed information about all records from the drive*)
	END_VAR
	VAR
		C_Axis : UDINT; (*internal variable*)
		IS : MC_0098_IS_TYP; (*internal structure*)
	END_VAR
END_FUNCTION_BLOCK

FUNCTION_BLOCK MC_BR_CyclicWrite (*enters a specified ParID in the cyclic data to drive*)
	VAR_INPUT
		Axis : UDINT; (*axis reference*)
		Enable : BOOL; (*specified ParID is written to the drive as long as enable is TRUE*)
		ParID : UINT; (*ParID which should be written to the drive*)
		DataAddress : UDINT; (*data address of the variable with the value for the ParID*)
		DataType : UINT; (*data type of the ParID*)
		Mode : UINT; (*currently not used*)
	END_VAR
	VAR_OUTPUT
		Valid : BOOL; (*when set the output is valid*)
		Busy : BOOL; (*function block is not finished*)
		Error : BOOL; (*error occurred in FB*)
		ErrorID : UINT; (*error number*)
	END_VAR
	VAR
		C_Axis : UDINT; (*internal variable*)
		IS : MC_0070_IS_TYP; (*internal variable*)
	END_VAR
END_FUNCTION_BLOCK

FUNCTION_BLOCK MC_BR_DigitalCamSwitch (*allows a digital output (Track) to be set whenever the axis is inside a position window*)
	VAR_INPUT
		Enable : BOOL; (*when set the FB parameters are downloaded*)
		Switches : MC_MASTER_SWITCHES_REF; (*reference to the switching actions*)
		OutputOptions : MC_OUTPUT_OPTIONS_REF; (*reference to the output options*)
		TrackOptions : MC_TRACK_OPTIONS_REF; (*reference to the track options*)
		SwitchSelector : USINT; (*selection of the switching data*)
		EnableValue : BOOL; (*enable the output of the state of the track on the FB output*)
		EnableParID : BOOL; (*enable the output of the state of the track on the specified ParID*)
		EnableDigOut : BOOL; (*enable the output of of the state of the track on a plug-in module*)
		ChangeSwitches : BOOL; (*change the active switching data*)
		InitSwitches : BOOL; (*initialize new switching parameters*)
		InitTrackOptions : BOOL; (*initialize new track options*)
	END_VAR
	VAR_OUTPUT
		InOperation : BOOL; (*is set after all parameters are transferred*)
		Busy : BOOL; (*the function block is active*)
		Error : BOOL; (*error occured in FB*)
		ErrorID : UINT; (*error number*)
		SwitchesChanged : BOOL; (*the active switching data has been changed*)
		SwitchesInitialized : BOOL; (*new switching parameters are initialized*)
		TrackOptionsInitialized : BOOL; (*new track options initialized*)
		Value : BOOL; (*actual state of the track*)
		ActualSwitches : USINT; (*actual active switches*)
	END_VAR
	VAR
		IS : MC_0107_IS_TYP; (*internal variable*)
		C_Master : UDINT; (*internal variable*)
		C_Slave : UDINT; (*internal variable*)
	END_VAR
END_FUNCTION_BLOCK

FUNCTION_BLOCK MC_BR_DownloadCamProfileObj (*transfers a cam profile object to the drive*)
	VAR_INPUT
		Axis : UDINT; (*axis reference*)
		Execute : BOOL; (*download camprofile at rising edge*)
		DataObjectName : STRING[12]; (*name of the data object*)
		Index : UINT; (*index for cam profile data object*)
		Periodic : BOOL; (*select if paeriodic or non periodic*)
	END_VAR
	VAR_OUTPUT
		Done : BOOL; (*download completed*)
		Busy : BOOL; (*function block is not finished*)
		Error : BOOL; (*error occurred in FB*)
		ErrorID : UINT; (*error number*)
	END_VAR
	VAR
		C_Axis : UDINT; (*internal variable*)
		C_DataObjectName : STRING[12]; (*internal variable*)
		LockIDPar : USINT; (*internal variable*)
		C_Error : BOOL; (*internal variable*)
		C_Index : UINT; (*internal variable*)
		C_ErrorID : UINT; (*internal variable*)
		C_Periodic : BOOL; (*internal variable*)
		C_Done : BOOL; (*internal variable*)
		state : USINT; (*internal variable*)
	END_VAR
END_FUNCTION_BLOCK

FUNCTION_BLOCK MC_BR_DownloadCamProfileData (*transfers cam profile data to the drive*)
	VAR_INPUT
		Axis : UDINT; (*axis reference*)
		Execute : BOOL; (*download cam profile at rising edge*)
		DataAddress : UDINT; (*address of cam profile data*)
		Index : UINT; (*index for cam profile data object*)
		Periodic : BOOL; (*decides if periodic or not*)
	END_VAR
	VAR_OUTPUT
		Done : BOOL; (*download completed*)
		Busy : BOOL; (*function block is not fnished*)
		Error : BOOL; (*error occurred in FB*)
		ErrorID : UINT; (*error number*)
	END_VAR
	VAR
		C_Axis : UDINT; (*internal variable*)
		C_DataAddress : UDINT; (*internal variable*)
		C_Index : UINT; (*internal variable*)
		C_ErrorID : UINT; (*internal variable*)
		C_Error : BOOL; (*internal variable*)
		C_Periodic : BOOL; (*internal variable*)
		C_Done : BOOL; (*internal variable*)
		state : USINT; (*internal variable*)
		LockIDPar : USINT; (*internal variable*)
	END_VAR
END_FUNCTION_BLOCK

FUNCTION_BLOCK MC_BR_DownloadParSequ (*downloads a parameter sequence*)
	VAR_INPUT
		Axis : UDINT; (*axis reference*)
		Execute : BOOL; (*download parameter sequence at rising edge*)
		DataAddress : UDINT; (*data address of the parameter sequence*)
	END_VAR
	VAR_OUTPUT
		Done : BOOL; (*download completed*)
		Busy : BOOL; (*function block is not finished*)
		Error : BOOL; (*error occurred*)
		ErrorID : UINT; (*error number*)
	END_VAR
	VAR
		Reserve1 : UINT; (*internal variable*)
		C_Axis : UDINT; (*internal variable*)
		C_DataAddress : UDINT; (*internal variable*)
		C_Done : BOOL; (*internal variable*)
		C_Error : BOOL; (*internal variable*)
		C_ErrorID : UINT; (*internal variable*)
		LockIDPar : USINT; (*internal variable*)
		Reserve2 : USINT; (*internal variable*)
		SizeOfFormat : UDINT; (*internal variable*)
		Reserve3 : UDINT; (*internal variable*)
		index : USINT; (*internal variable*)
		state : USINT; (*internal variable*)
	END_VAR
END_FUNCTION_BLOCK

FUNCTION_BLOCK MC_BR_EventMoveAbsolute (*starts an absolute positioning on the drive after a specified event*)
	VAR_INPUT
		Axis : UDINT; (*axis reference*)
		Execute : BOOL; (*wait for the event at rising edge*)
		EventInput : MC_BR_EVINPUT_REF; (*input that is used as event source*)
		Position : REAL; (*target position for the movement*)
		Velocity : REAL; (*maximum velocity*)
		Acceleration : REAL; (*maximum acceleration*)
		Deceleration : REAL; (*maximum deceleration*)
		Direction : USINT; (*direction of movement*)
		Mode : UINT; (*mcONCE or mcCYCLIC or mcCYCLIC_ALL_EVENTS*)
		PositionParID : UINT; (*ParID from which the target position is read*)
	END_VAR
	VAR_OUTPUT
		InPosition : BOOL; (*target position reached*)
		Busy : BOOL; (*function block is not finished*)
		CommandAborted : BOOL; (*function block aborted by another command*)
		Error : BOOL; (*error occurred in FB*)
		ErrorID : UINT; (*error number*)
		WaitingForEvent : BOOL; (*waiting for event*)
	END_VAR
	VAR
		C_Axis : UDINT; (*internal variable*)
		C_EventInput : MC_BR_EVINPUT_REF; (*internal variable*)
		C_Execute : BOOL; (*internal variable*)
		C_Position : DINT; (*internal variable*)
		C_Velocity : REAL; (*internal variable*)
		C_Acceleration : REAL; (*internal variable*)
		C_Deceleration : REAL; (*internal variable*)
		C_Mode : UINT; (*internal variable*)
		C_PositionParID : UINT; (*internal variable*)
		C_InPosition : BOOL; (*internal variable*)
		C_WaitingForEvent : BOOL; (*internal variable*)
		C_Busy : BOOL; (*internal variable*)
		C_CommandAborted : BOOL; (*internal variable*)
        C_ErrorID : UINT; (*internal variable*)
        C_Error : BOOL; (*internal variable*)
        C_Direction : USINT; (*internal variable*)
		C_CommandedOffset : DINT; (*internal variable*)
		CmpIndex : UINT; (*internal variable*)
		VarIndex : UINT; (*internal variable*)
		EvMoveStatusOffset : UINT; (*internal variable*)
		EvMoveStatusRecIndex : USINT; (*internal variable*)
		SavedFrDrvCnt : USINT; (*internal variable*)
		WaitEvMoveStatusValid : BOOL; (*internal variable*)
		C_MoveActive : BOOL; (*internal variable*)
		state : USINT; (*internal variable*)
		LockID : USINT; (*internal variable*)
		LockIDPar : USINT; (*internal variable*)
		MoveID : USINT; (*internal variable*)
		WaitForTelegrams : BOOL; (*internal variable*)
        oldMoveID : USINT; (*internal variable*)
	END_VAR
END_FUNCTION_BLOCK

FUNCTION_BLOCK MC_BR_EventMoveAdditive (*starts a movement on the drive by a set distance after a specified event*)
	VAR_INPUT
		Axis : UDINT; (*axis reference*)
		Execute : BOOL; (*wait for the event at rising edge*)
		EventInput : MC_BR_EVINPUT_REF; (*input that is used as event source*)
		Distance : REAL; (*relative distance of the movement*)
		Velocity : REAL; (*maximum velocity*)
		Acceleration : REAL; (*maximum acceleration*)
		Deceleration : REAL; (*maximum deceleration*)
		Mode : UINT; (*mcONCE or mcCYCLIC or mcCYCLIC_ALL_EVENTS*)
		DistanceParID : UINT; (*ParID from which the distance is read*)
	END_VAR
	VAR_OUTPUT
		InPosition : BOOL; (*target position reached*)
		Busy : BOOL; (*function block is not finished*)
		CommandAborted : BOOL; (*function block aborted by another command*)
		Error : BOOL; (*error occurred in FB*)
		ErrorID : UINT; (*error number*)
		WaitingForEvent : BOOL; (*waiting for the event*)
	END_VAR
	VAR
		C_Axis : UDINT; (*internal variable*)
		C_EventInput : MC_BR_EVINPUT_REF; (*internal variable*)
		C_Execute : BOOL; (*internal variable*)
		C_Distance : DINT; (*internal variable*)
		C_Velocity : REAL; (*internal variable*)
		C_Acceleration : REAL; (*internal variable*)
		C_Deceleration : REAL; (*internal variable*)
		C_Mode : UINT; (*internal variable*)
		C_DistanceParID : UINT; (*internal variable*)
		C_InPosition : BOOL; (*internal variable*)
		C_WaitingForEvent : BOOL; (*internal variable*)
		C_Busy : BOOL; (*internal variable*)
		C_CommandAborted : BOOL; (*internal variable*)
        C_ErrorID : UINT; (*internal variable*)
        C_Error : BOOL; (*internal variable*)
        Reserve : USINT; (*internal variable*)
		C_CommandedOffset : DINT; (*internal variable*)
		C_CommandedPosition : DINT; (*internal variable*)
		CmpIndex : UINT; (*internal variable*)
		VarIndex : UINT; (*internal variable*)
		EvMoveStatusOffset : UINT; (*internal variable*)
		EvMoveStatusRecIndex : USINT; (*internal variable*)
		SavedFrDrvCnt : USINT; (*internal variable*)
		WaitEvMoveStatusValid : BOOL; (*internal variable*)
		C_MoveActive : BOOL; (*internal variable*)
		state : USINT; (*internal variable*)
		LockID : USINT; (*internal variable*)
		LockIDPar : USINT; (*internal variable*)
		MoveID : USINT; (*internal variable*)
        WaitForTelegrams : BOOL; (*internal variable*)
        oldMoveID : USINT; (*internal variable*)
	END_VAR
END_FUNCTION_BLOCK

FUNCTION_BLOCK MC_BR_EventMoveVelocity (*starts a controlled movement with a specified velocity after a specified event*)
	VAR_INPUT
		Axis : UDINT; (*axis reference*)
		Execute : BOOL; (*wait for the event at rising edge*)
		EventInput : MC_BR_EVINPUT_REF; (*input that is used as event source*)
		Velocity : REAL; (*target velocity*)
		Acceleration : REAL; (*maximum acceleration*)
		Deceleration : REAL; (*maximum deceleration*)
		Direction : USINT; (*direction of movement*)
		Mode : UINT; (*mcONCE or mcCYCLIC_ALL_EVENTS*)
		VelocityParID : UINT; (*ParID from which the velocity is read*)
	END_VAR
	VAR_OUTPUT
		InVelocity : BOOL; (*specified velocity achieved*)
		Busy : BOOL; (*function block is not finished*)
		CommandAborted : BOOL; (*function block aborted by another command*)
		Error : BOOL; (*error occurred in FB*)
		ErrorID : UINT; (*error number*)
		WaitingForEvent : BOOL; (*waiting for the event*)
	END_VAR
	VAR
		C_Axis : UDINT; (*internal variable*)
		C_Execute : BOOL; (*internal variable*)
		C_EventInput : MC_BR_EVINPUT_REF; (*internal variable*)
		C_Velocity : REAL; (*internal variable*)
		C_Acceleration : REAL; (*internal variable*)
		C_Deceleration : REAL; (*internal variable*)
		C_Direction : USINT; (*internal variable*)
		LockID : USINT; (*internal variable*)
		LockIDPar : USINT; (*internal variable*)
		C_Mode : UINT; (*internal variable*)
		C_VelocityParID : UINT; (*internal variable*)
		C_InVelocity : BOOL; (*internal variable*)
		C_WaitingForEvent : BOOL; (*internal variable*)
		C_Busy : BOOL; (*internal variable*)
		C_CommandAborted : BOOL; (*internal variable*)
		C_Error : BOOL; (*internal variable*)
		C_ErrorID : UINT; (*internal variable*)
		CmpIndex : UINT; (*internal variable*)
		VarIndex : UINT; (*internal variable*)
		EvMoveStatusOffset : UINT; (*internal variable*)
		EvMoveStatusRecIndex : USINT; (*internal variable*)
		Reserve1 : USINT; (*internal variable*)
		VelocityOffset : UINT; (*internal variable*)
		VelocityRecIndex : USINT; (*internal variable*)
		SavedFrDrvCnt : USINT; (*internal variable*)
		WaitEvMoveStatusValid : BOOL; (*internal variable*)
		C_MoveActive : BOOL; (*internal variable*)
		state : USINT; (*internal variable*)
		MoveID : USINT; (*internal variable*)
		WaitForTelegrams : BOOL; (*internal variable*)
	END_VAR
END_FUNCTION_BLOCK

FUNCTION_BLOCK MC_BR_GearIn (*commands a ratio between the velocity of the master and slave axes*)
	VAR_INPUT
		Master : UDINT; (*axis reference of the master axis *)
		Slave : UDINT; (*axis reference of the slave axis *)
		Enable : BOOL; (*the gear ratio is active as long as this input is set*)
		InitData : BOOL; (*starts transferring the parameters*)
		RatioNumerator : DINT; (*gear ratio numerator*)
		RatioDenominator : DINT; (*gear ratio denominator*)
		AdvancedParameters : MC_ADVANCED_GEAR_PAR_REF; (*additional inputs for advanced usage of FB*)
	END_VAR
	VAR_OUTPUT
		Active : BOOL; (*parameters are transferred and FB is active*)
		Busy : BOOL; (*function block is enabled *)
		CommandAborted : BOOL; (*function block aborted by another FB*)
		Error : BOOL; (*error occured in FB*)
		ErrorID : UINT; (*error number*)
		DataInitialized : BOOL; (*transferring parameters is completed *)
		InGear : BOOL; (*commanded gear ratio reached*)
	END_VAR
	VAR
		C_Master : UDINT; (*internal variable*)
		C_Slave : UDINT; (*internal variable*)
		IS : MC_0126_IS_TYP; (*internal variable*)
	END_VAR
END_FUNCTION_BLOCK

FUNCTION_BLOCK MC_BR_GetCamMasterPosition (*get the master position according to cam profile and slave position*)
	VAR_INPUT
		Master : UDINT; (*master axis reference*)
		Slave : UDINT; (*slave axis reference*)
		Execute : BOOL; (*start master position determination*)
		DataObjectName : STRING[12]; (*name of cam profile data object*)
		DataAddress : UDINT; (*address of cam profile data*)
		MasterStartPosition : REAL; (*master position within cam to start determination of slave position*)
		SlavePosition : REAL; (*slave position within cam to determine master position*)
		MasterFactor : UDINT; (*multiplication factor of the cam on the master axis*)
		SlaveFactor : DINT; (*multiplication factor of the cam on the slave axis*)
	END_VAR
	VAR_OUTPUT
		Done : BOOL; (*master position determination finished*)
		Busy : BOOL; (*function block is not finished*)
		Error : BOOL; (*error occurred in FB*)
		ErrorID : UINT; (*error number*)
		MasterPosition : REAL; (*determined master position*)
	END_VAR
	VAR
		C_Master : UDINT; (*internal variable*)
		C_Slave : UDINT; (*internal variable*)
		IS : MC_0084_IS_TYP; (*internal variable*)
	END_VAR
END_FUNCTION_BLOCK

FUNCTION_BLOCK MC_BR_GetCamSlavePosition (*get the slave position according to cam profile and master position*)
	VAR_INPUT
		Master : UDINT; (*master axis reference*)
		Slave : UDINT; (*slave axis reference*)
		Execute : BOOL; (*start slave position determination*)
		DataObjectName : STRING[12]; (*name of cam profile data object*)
		DataAddress : UDINT; (*address of cam profile data*)
		MasterPosition : REAL; (*master position within cam to determine slave position*)
		MasterFactor : UDINT; (*multiplication factor of the cam on the master axis*)
		SlaveFactor : DINT; (*multiplication factor of the cam on the slave axis*)
	END_VAR
	VAR_OUTPUT
		Done : BOOL; (*slave position determination finished*)
		Busy : BOOL; (*function block is not finished*)
		Error : BOOL; (*error occurred in FB*)
		ErrorID : UINT; (*error number*)
		SlavePosition : REAL; (*determined slave position*)
	END_VAR
	VAR
		C_Master : UDINT; (*internal variable*)
		C_Slave : UDINT; (*internal variable*)
		IS : MC_0083_IS_TYP; (*internal variable*)
	END_VAR
END_FUNCTION_BLOCK

FUNCTION_BLOCK MC_BR_GetErrorText (*determines the error text for an error record*)
	VAR_INPUT
		Execute : BOOL; (*error text determined after a rising edge*)
		Configuration : MC_ERRORTEXTCONFIG_REF; (*FB configuration*)
		ErrorRecord : MC_ERRORRECORD_REF; (*error record for which the error text should be determined*)
	END_VAR
	VAR_OUTPUT
		Done : BOOL; (*error text determined*)
		Busy : BOOL; (*function block is not finished*)
		Error : BOOL; (*error occurred in FB*)
		ErrorID : UINT; (*error number*)
	END_VAR
	VAR
		IS : MC_0077_IS_TYP; (*internal variable*)
	END_VAR
END_FUNCTION_BLOCK

FUNCTION_BLOCK MC_BR_GetHardwareInfo (*determines hardware information of drive components*)
	VAR_INPUT
		Axis : UDINT; (*axis reference*)
		Execute : BOOL; (*determine ParID information at rising edge*)
	END_VAR
	VAR_OUTPUT
		Done : BOOL; (*command executed*)
		Busy : BOOL; (*function block is not finished*)
		Error : BOOL; (*error occurred in FB*)
		ErrorID : UINT; (*error number*)
		HardwareInfo : MC_HARDWARE_INFO_REF; (*hardware information of drive components*)
	END_VAR
	VAR
		C_Axis : UDINT; (*internal variable*)
		IS : MC_0109_IS_TYP; (*intern variable*)
	END_VAR
END_FUNCTION_BLOCK

FUNCTION_BLOCK MC_BR_GetParIDTransferInfo (*determines ParID transfer information of an axis*)
	VAR_INPUT
		Axis : UDINT; (*axis reference*)
		Execute : BOOL; (*determine ParID transfer information at rising edge*)
	END_VAR
	VAR_OUTPUT
		Done : BOOL; (*command executed*)
		Busy : BOOL; (*function block is not finished*)
		Error : BOOL; (*error occurred in FB*)
		ErrorID : UINT; (*error number*)
		FreeSendChannels : USINT; (*number of free send channels on the axis*)
		FreeReceiveChannels : USINT; (*number of free receive channels on the axis*)
		ParIDTransferInfo : MC_TRANSFER_INFO_REF; (*ParID transfer information of the axis*)
	END_VAR
	VAR
		C_Axis : UDINT; (*internal variable*)
		IS : MC_0121_IS_TYP; (*intern variable*)
	END_VAR
END_FUNCTION_BLOCK

FUNCTION_BLOCK MC_BR_HomeAcpEncoder (*homes an external encoder*)
	VAR_INPUT
		AcpEncoder : MC_ACP_ENCOD_REF; (*ACOPOS encoder*)
		Execute : BOOL; (*starts homing the encoder*)
		HomingParameters : MC_ACP_ENCOD_PARAM_REF; (*parameter for homing the encoder*)
	END_VAR
	VAR_OUTPUT
		Done : BOOL; (*homing procedur is completed*)
		Busy : BOOL; (*function block is not finished*)
		CommandAborted : BOOL; (*function block aborted by another command*)
		Error : BOOL; (*error occurred in FB*)
		ErrorID : UINT; (*error number*)
		EncoderOffset : DINT; (*home offset after homing procedur*)
	END_VAR
	VAR
		C_Axis : UDINT; (*internal variable*)
		IS : MC_0068_IS_TYP; (*internal variable*)
	END_VAR
END_FUNCTION_BLOCK

FUNCTION_BLOCK MC_BR_InitAutData (*initialize the parameters of cam profile automat*)
	VAR_INPUT
		Slave : UDINT; (*slave axis*)
		Execute : BOOL; (*starts initialization at rising edge*)
		InitOptions : MC_AUTINITOPTIONS_REF; (*configuration of the FB*)
		AdrAutData : UDINT; (*address of the automat data structure*)
	END_VAR
	VAR_OUTPUT
		Done : BOOL; (*initialization complete*)
		Busy : BOOL; (*initialization active*)
		Error : BOOL; (*error occurred in FB*)
		ErrorID : UINT; (*error number*)
	END_VAR
	VAR
		C_Master : UDINT; (*internal variable*)
		C_Slave : UDINT; (*internal variable*)
		IS : MC_0076_IS_TYP; (*internal variable*)
	END_VAR
END_FUNCTION_BLOCK

FUNCTION_BLOCK MC_BR_InitAutEvent (*initializes the parameters of an event for the specified cam automat state*)
	VAR_INPUT
		Slave : UDINT; (*axis reference of the slave axis*)
		Execute : BOOL; (*initialize parameter at rising edge*)
		StateIndex : USINT; (*state index for this event*)
		EventIndex : USINT; (*index for parameter set for an event*)
		Type : USINT; (*event type*)
		Attribute : USINT; (*event attribute*)
		Action : UDINT; (*action at state transition*)
		NextState : USINT; (*index for the next state*)
	END_VAR
	VAR_OUTPUT
		Done : BOOL; (*automat event initialized*)
		Busy : BOOL; (*function block is not finished*)
		Error : BOOL; (*error occurred in FB*)
		ErrorID : UINT; (*error number*)
	END_VAR
	VAR
		C_Slave : UDINT; (*internal variable*)
		C_Execute : BOOL; (*internal variable*)
		C_StateIndex : USINT; (*internal variable*)
		C_EventIndex : USINT; (*internal variable*)
		C_Type : USINT; (*internal variable*)
		C_Attribute : USINT; (*internal variable*)
		C_Action : UDINT; (*internal variable*)
		C_NextState : USINT; (*internal variable*)
		LockIDPar : USINT; (*internal variable*)
		C_Done : BOOL; (*internal variable*)
		C_Error : BOOL; (*internal variable*)
		C_ErrorID : UINT; (*internal variable*)
		Reserve : UDINT; (*internal variable*)
		state : USINT; (*internal variable*)
	END_VAR
END_FUNCTION_BLOCK

FUNCTION_BLOCK MC_BR_InitAutPar (*initializes the general parameters of the cam automat*)
	VAR_INPUT
		Master : UDINT; (*axis reference of the master axis*)
		Slave : UDINT; (*axis reference of the slave axis*)
		Execute : BOOL; (*initialize parameter at rising edge*)
		StartPosition : REAL; (*start position of the master axis*)
		StartInterval : REAL; (*start interval for the master axis*)
		StartState : USINT; (*index for the start state*)
		StartMaRelPos : REAL; (*relative master position in the cam profile*)
		MaxMasterVelocity : REAL; (*maximum speed of the master axis*)
		MasterParID : UINT; (*use this ParID from the master axis instead of the set position*)
		AddMasterParID : UINT; (*ParID of the additive master axis*)
		AddSlaveParID : UINT; (*ParID of the additive slave axis*)
		SlaveFactorParID : UINT; (*ParID for multiplication factor of the slave axis*)
		EventParID : UINT; (*ParID for event input*)
		SlaveLatchParID : UINT; (*ParID for the latch value of the slave axis*)
	END_VAR
	VAR_OUTPUT
		Done : BOOL; (*automat parameters initialized*)
		Busy : BOOL; (*function block not finished*)
		Error : BOOL; (*error occurred in FB*)
		ErrorID : UINT; (*error number*)
	END_VAR
	VAR
		Reserve1 : USINT; (*internal variable*)
		LockIDReceive : USINT; (*internal variable*)
		C_Master : UDINT; (*internal variable*)
		C_Slave : UDINT; (*internal variable*)
		C_Execute : BOOL; (*internal variable*)
		C_StartPosition : DINT; (*internal variable*)
		C_StartInterval : DINT; (*internal variable*)
		C_StartState : USINT; (*internal variable*)
		LockIDMa : USINT; (*internal variable*)
		LockIDPar : USINT; (*internal variable*)
		LockIDSend : USINT; (*internal variable*)
		C_StartMaRelPos : DINT; (*internal variable*)
		C_MaxMasterVelocity : REAL; (*internal variable*)
		Reserve2 : UDINT; (*internal variable*)
		C_MasterParID : UINT; (*internal variable*)
		C_AddMasterParID : UINT; (*internal variable*)
		C_AddSlaveParID : UINT; (*internal variable*)
		C_SlaveFactorParID : UINT; (*internal variable*)
		C_EventParID : UINT; (*internal variable*)
		C_SlaveLatchParID : UINT; (*internal variable*)
		C_Done : BOOL; (*internal variable*)
		C_Error : BOOL; (*internal variable*)
		C_ErrorID : UINT; (*internal variable*)
		sendSlot : USINT; (*internal variable*)
		readSlot : USINT; (*internal variable*)
		state : USINT; (*internal variable*)
	END_VAR
END_FUNCTION_BLOCK

FUNCTION_BLOCK MC_BR_InitAutState (*initializes the parameters of a cam automat state*)
	VAR_INPUT
		Master : UDINT; (*axis reference of the master axis*)
		Slave : UDINT; (*axis reference of the slave axis*)
		Execute : BOOL; (*initialize parameter at rising edge*)
		StateIndex : USINT; (*index of a parameter set for a state*)
		CamProfileIndex : UINT; (*index of cam profile data for one state*)
		MasterFactor : UDINT; (*multiplication factor for the master axis*)
		SlaveFactor : DINT; (*multiplication factor for the slave axis*)
		RepeatCounterInit : UINT; (*start value state repeats for the ncCOUNT event*)
		RepeatCounterSet : UINT; (*counter state repeats for the ncCOUNT event*)
		CompMode : USINT; (*compensation gear mode*)
		MasterCompDistance : REAL; (*compensation distance for the master axis*)
		SlaveCompDistance : REAL; (*compensation distance for the slave axis*)
		ExtendedCompLimits : USINT; (*extended compensation limits*)
		MinMasterCompDistance : REAL; (*minimum compensation distance for the master axis*)
		MinSlaveCompDistance : REAL; (*minimum compensation distance for the slave axis*)
		MaxSlaveCompDistance : REAL; (*maximum compensation distance for the slave axis*)
		MinSlaveCompVelocity : REAL; (*minimum speed of the slave axis in the compensation*)
		MaxSlaveCompVelocity : REAL; (*maximum speed of the slave axis in the compensation*)
		MaxSlaveAccelComp1 : REAL; (*maximum acceleration of the slave axis in compensation phase 1*)
		MaxSlaveAccelComp2 : REAL; (*maximum acceleration of the slave axis in compensation phase 2*)
		SlaveCompJoltTime : REAL; (*jolt time of the slave axis in the compensation*)
		MasterParID : UINT; (*master ParID for this state*)
	END_VAR
	VAR_OUTPUT
		Done : BOOL; (*automat state parameters initialized*)
		Busy : BOOL; (*function block is not finished*)
		Error : BOOL; (*error occurred in FB*)
		ErrorID : UINT; (*error number*)
	END_VAR
	VAR
		C_Master : UDINT; (*internal variable*)
		C_Slave : UDINT; (*internal variable*)
		C_Execute : BOOL; (*internal variable*)
		C_StateIndex : USINT; (*internal variable*)
		Reserve1 : USINT; (*internal variable*)
		C_CamProfileIndex : UINT; (*internal variable*)
		C_MasterFactor : DINT; (*internal variable*)
		C_SlaveFactor : DINT; (*internal variable*)
		C_RepeatCounterInit : UINT; (*internal variable*)
		Reserve2 : UINT; (*internal variable*)
		C_RepeatCounterSet : UINT; (*internal variable*)
		C_CompMode : USINT; (*internal variable*)
		LockIDPar : USINT; (*internal variable*)
		C_MasterCompDistance : DINT; (*internal variable*)
		C_SlaveCompDistance : DINT; (*internal variable*)
		C_ExtendedCompLimits : USINT; (*internal variable*)
		Reserve3 : USINT; (*internal variable*)
		Reserve4 : UINT; (*internal variable*)
		C_MinMasterCompDistance : DINT; (*internal variable*)
		C_MinSlaveCompDistance : DINT; (*internal variable*)
		C_MaxSlaveCompDistance : DINT; (*internal variable*)
		C_MinSlaveCompVelocity : REAL; (*internal variable*)
		C_MaxSlaveCompVelocity : REAL; (*internal variable*)
		C_MaxSlaveAccelComp1 : REAL; (*internal variable*)
		C_MaxSlaveAccelComp2 : REAL; (*internal variable*)
		C_SlaveCompJoltTime : REAL; (*internal variable*)
		C_MasterParID : UINT; (*internal variable*)
		C_Done : BOOL; (*internal variable*)
		C_Error : BOOL; (*internal variable*)
		C_ErrorID : UINT; (*internal variable*)
		Reserve5 : UDINT; (*internal variable*)
		state : USINT; (*internal variable*)
	END_VAR
END_FUNCTION_BLOCK

FUNCTION_BLOCK MC_BR_InitAxisPar (*initializes the axis parameter in the axis data structure*)
	VAR_INPUT
		Axis : UDINT; (*axis reference*)
		Execute : BOOL; (*initializes the axis parameter at rising edge*)
	END_VAR
	VAR_OUTPUT
		Done : BOOL; (*initialization of the data is finished*)
		Busy : BOOL; (*function block is not finished*)
		Error : BOOL; (*error occurred in FB*)
		ErrorID : UINT; (*error number*)
	END_VAR
	VAR
		C_Axis : UDINT; (*internal variable*)
		state : USINT; (*internal variable*)
		LockIDPar : USINT; (*internal variable*)
		C_ErrorID : UINT; (*internal variable*)
		C_Error : BOOL; (*internal variable*)
		pInit : REFERENCE TO USINT; (*internal variable*)
		pError : REFERENCE TO USINT; (*internal variable*)
	END_VAR
END_FUNCTION_BLOCK

FUNCTION_BLOCK MC_BR_InitAxisSubjectPar (*enables the user to selectively initialize structure elements from the axis data structure*)
	VAR_INPUT
		Axis : UDINT; (*axis reference*)
		Execute : BOOL; (*initializes the axis parameters in the selected axis structure*)
		Subject : UINT; (*subject of the axis structure whose data should be initialized*)
	END_VAR
	VAR_OUTPUT
		Done : BOOL; (*initialization of the data finished*)
		Busy : BOOL; (*function block is not finished*)
		Error : BOOL; (*error occurred in function block*)
		ErrorID : UINT; (*error number*)
	END_VAR
	VAR
		C_Axis : UDINT; (*internal variable*)
		C_Subject : UINT; (*internal variable*)
		C_ErrorID : UINT; (*internal varaible*)
		C_Error : BOOL; (*internal variable*)
		state : USINT; (*internal variable*)
		LockIDPar : USINT; (*internal variable*)
		pInit : REFERENCE TO USINT; (*internal variable*)
		pError : REFERENCE TO USINT; (*internal variable*)
		CheckModeBits : UDINT; (*internal variable*)
	END_VAR
END_FUNCTION_BLOCK

FUNCTION_BLOCK MC_BR_InitCyclicRead (*adds the specified ParID to the cyclic data from drive*)
	VAR_INPUT
		Axis : UDINT; (*axis refrence*)
		Execute : BOOL; (*initialize cyclic data read at rising edge*)
		ParID : UINT; (*number of the parameter ID to read cyclically*)
		DataAddress : UDINT; (*address of the user variable*)
		DataType : UINT; (*data type of user variable*)
		Mode : UINT; (*currently not used*)
	END_VAR
	VAR_OUTPUT
		Done : BOOL; (*requested parameter is available*)
		Busy : BOOL; (*function block is not finished*)
		Error : BOOL; (*error occurred in FB*)
		ErrorID : UINT; (*error number*)
	END_VAR
	VAR
		LockID : USINT; (*internal variable*)
		LockIDPar : USINT; (*internal variable*)
		C_Axis : UDINT; (*internal variable*)
		C_Execute : BOOL; (*internal variable*)
		C_ParID : UINT; (*internal variable*)
		Reserve1 : UINT; (*internal variable*)
		C_DataAddress : UDINT; (*internal variable*)
		C_DataType : UINT; (*internal variable*)
		C_Mode : UINT; (*internal variable*)
		C_Done : BOOL; (*internal variable*)
		C_Error : BOOL; (*internal variable*)
		C_ErrorID : UINT; (*internal variable*)
		ParIDOffset : UINT; (*internal variable*)
		Reserve2 : UDINT; (*internal variable*)
		Reserve3 : USINT; (*internal variable*)
		ParIDRecIndex : USINT; (*internal variable*)
		Reserve4 : USINT; (*internal variable*)
		DataLength : USINT; (*internal variable*)
		state : USINT; (*internal variable*)
	END_VAR
END_FUNCTION_BLOCK

FUNCTION_BLOCK MC_BR_InitCyclicWrite (*adds the specified ParID to the cyclic data to the drive*)
	VAR_INPUT
		Axis : UDINT; (*axis reference*)
		Execute : BOOL; (*initialize cyclic data write at rising edge*)
		ParID : UINT; (*number of the Parameter ID to write cyclically*)
		DataAddress : UDINT; (*address of the user variable*)
		DataType : UINT; (*data type of the user variable*)
		Mode : UINT; (*currently not used*)
	END_VAR
	VAR_OUTPUT
		Done : BOOL; (*initialization of the data write command is done*)
		Busy : BOOL; (*function block is not finished*)
		Error : BOOL; (*error occurred in FB*)
		ErrorID : UINT; (*error number*)
	END_VAR
	VAR
		LockID : USINT; (*internal variable*)
		LockIDPar : USINT; (*internal variable*)
		C_Axis : UDINT; (*internal variable*)
		C_Execute : BOOL; (*internal variable*)
		C_ParID : UINT; (*internal variable*)
		Reserve1 : UINT; (*internal variable*)
		C_DataAddress : UDINT; (*internal variable*)
		C_DataType : UINT; (*internal variable*)
		C_Mode : UINT; (*internal variable*)
		Reserve2 : UDINT; (*internal variable*)
		C_Done : BOOL; (*internal variable*)
		C_Error : BOOL; (*internal variable*)
		C_ErrorID : UINT; (*internal variable*)
		ParIDParIndex : USINT; (*internal variable*)
		DataLength : USINT; (*internal variable*)
		state : USINT; (*internal variable*)
	END_VAR
END_FUNCTION_BLOCK

FUNCTION_BLOCK MC_BR_InitEndlessPosition (*initialize memory for endless position storage*)
	VAR_INPUT
		Axis : UDINT; (*axis reference*)
		Execute : BOOL; (*initialize memory storage at rising edge*)
		DataAddress : UDINT; (*data address of momory storage for endless position*)
	END_VAR
	VAR_OUTPUT
		Done : BOOL; (*memory storage for endless position was initialized*)
		Busy : BOOL; (*function block is not finished*)
		Error : BOOL; (*error occurred in FB*)
		ErrorID : UINT; (*error number*)
	END_VAR
	VAR
		C_Axis : UDINT; (*internal variable*)
		C_ErrorID : UINT; (*internal variable*)
		C_Error : BOOL; (*internal variable*)
		state : USINT; (*internal variable*)
	END_VAR
END_FUNCTION_BLOCK

FUNCTION_BLOCK MC_BR_InitEndlessPosAcpEnc (*initialize memory for endless position storage for external encoder*)
	VAR_INPUT
		AcpEncoder : MC_ACP_ENCOD_REF; (*ACOPOS encoder*)
		Execute : BOOL; (*initialize memory storage at rising edge*)
		DataAddress : UDINT; (*data address of memory storage for endless position*)
	END_VAR
	VAR_OUTPUT
		Done : BOOL; (*memory storage for endless position was initialized*)
		Busy : BOOL; (*function block is not finished*)
		Error : BOOL; (*error occurred in FB*)
		ErrorID : UINT; (*error number*)
		DataValid : BOOL; (*axis position can be restored from the endless position data*)
	END_VAR
	VAR
		C_Axis : UDINT; (*internal variable*)
		IS : MC_0138_IS_TYP; (*internal variable*)
	END_VAR
END_FUNCTION_BLOCK

FUNCTION_BLOCK MC_BR_InitMasterParIDTransfer (*initializes a cyclic ParID transfer from master to slave*)
	VAR_INPUT
		Master : UDINT; (*axis reference of the master axis*)
		Slave : UDINT; (*axis reference of the slave axis*)
		Execute : BOOL; (*initialize transfer at rising edge*)
		MasterParID : UINT; (*use this ParID from the master axis instead of the set position*)
		SlaveChannel : USINT; (*choose a slave channel*)
	END_VAR
	VAR_OUTPUT
		Done : BOOL; (*parameter transfer initialized*)
		Busy : BOOL; (*function block is not finished*)
		Error : BOOL; (*error occurred in FB*)
		ErrorID : UINT; (*error number*)
		ReceiveParID : UINT; (*ParID on Slave axis to use as master ParID*)
	END_VAR
	VAR
		C_Master : UDINT; (*internal variable*)
		C_Slave : UDINT; (*internal variable*)
		Reserve1 : UINT; (*internal variable*)
		Reserve2 : USINT; (*internal variable*)
		LockIDReceive : USINT; (*internal variable*)
		C_Execute : BOOL; (*internal variable*)
		C_MasterParID : UINT; (*internal variable*)
		C_SlaveChannel : USINT; (*internal variable*)
		C_Done : BOOL; (*internal variable*)
		C_Error : BOOL; (*internal variable*)
		LockIDSend : USINT; (*internal variable*)
		C_ErrorID : UINT; (*internal variable*)
		C_ReceiveParID : UINT; (*internal variable*)
		sendSlot : USINT; (*internal variable*)
		readSlot : USINT; (*internal variable*)
		state : USINT; (*internal variable*)
		LockIDMa : USINT; (*internal variable*)
		LockIDPar : USINT; (*internal variable*)
	END_VAR
END_FUNCTION_BLOCK

FUNCTION_BLOCK MC_BR_InitModPos (*initializes the modulo position parameters*)
	VAR_INPUT
		Axis : UDINT; (*axis reference*)
		Execute : BOOL; (*initialize the modulo position parameter with rising edge*)
		Period : UDINT; (*axis period*)
		Factor : UDINT; (*factor for conversion into init parameter module units*)
	END_VAR
	VAR_OUTPUT
		Done : BOOL; (*modulo position parameters were initialized*)
		Busy : BOOL; (*function block is not finished*)
		Error : BOOL; (*error occurred in FB*)
		ErrorID : UINT; (*error number*)
	END_VAR
	VAR
		C_Axis : UDINT; (*internal variable*)
		C_Period : UDINT; (*internal variable*)
		C_Factor : UDINT; (*internal variable*)
		C_ErrorID : UINT; (*internal varaible*)
		C_Error : BOOL; (*internal variable*)
		state : USINT; (*internal variable*)
		LockIDPar : USINT; (*internal variable*)
		C_Execute : BOOL; (*internal variable*)
	END_VAR
END_FUNCTION_BLOCK

FUNCTION_BLOCK MC_BR_InitParList (*initializes a parameter list*)
	VAR_INPUT
		Axis : UDINT; (*axis reference*)
		Execute : BOOL; (*initialize parameter list at rising edge*)
		DataAddress : UDINT; (*address of the parameter list*)
	END_VAR
	VAR_OUTPUT
		Done : BOOL; (*init completed*)
		Busy : BOOL; (*function block is not finished*)
		Error : BOOL; (*error occurred in FB*)
		ErrorID : UINT; (*error number*)
	END_VAR
	VAR
		LockIDPar : USINT; (*internal variable*)
		C_Error : BOOL; (*internal variable*)
		C_ErrorID : UINT; (*internal variable*)
		C_Axis : UDINT; (*internal variable*)
		C_DataAddress : UDINT; (*internal variable*)
		C_Done : BOOL; (*internal variable*)
		state : USINT; (*internal variable*)
	END_VAR
END_FUNCTION_BLOCK

FUNCTION_BLOCK MC_BR_InitParSequ (*initializes a parameter sequence*)
	VAR_INPUT
		Axis : UDINT; (*axis reference*)
		Execute : BOOL; (*initialize parameter sequence at rising edge*)
		DataAddress : UDINT; (*address of the parameter sequence*)
	END_VAR
	VAR_OUTPUT
		Done : BOOL; (*init completed*)
		Busy : BOOL; (*function block is not finished*)
		Error : BOOL; (*error occurred in FB*)
		ErrorID : UINT; (*error number*)
	END_VAR
	VAR
		C_Axis : UDINT; (*internal variable*)
		C_DataAddress : UDINT; (*internal variable*)
		Reserve1 : UINT; (*internal variable*)
		Reserve2 : UDINT; (*internal variable*)
		C_Error : BOOL; (*internal variable*)
		C_ErrorID : UINT; (*internal variable*)
		Reserve3 : UDINT; (*internal variable*)
		index : USINT; (*internal variable*)
		Reserve4 : UINT; (*internal variable*)
		state : USINT; (*internal variable*)
		LockIDPar : USINT; (*internal variable*)
	END_VAR
END_FUNCTION_BLOCK

FUNCTION_BLOCK MC_BR_InitParTabObj (*transfers and initializes the parameters contained in "DataObjName" on the specified axis*)
	VAR_INPUT
		Axis : UDINT; (*axis reference*)
		Execute : BOOL; (*initialize parameter table at rising edge*)
		DataObjectName : STRING[12]; (*name of the data object*)
	END_VAR
	VAR_OUTPUT
		Done : BOOL; (*initialization completed*)
		Busy : BOOL; (*function block is not finished*)
		Error : BOOL; (*error occurred in FB*)
		ErrorID : UINT; (*error number*)
	END_VAR
	VAR
		C_Axis : UDINT; (*internal variable*)
		C_DataObjectName : STRING[12]; (*internal variable*)
		C_ErrorID : UINT; (*internal variable*)
		C_Error : BOOL; (*internal variable*)
		C_Done : BOOL; (*internal variable*)
		LockIDPar : USINT; (*internal variable*)
		state : USINT; (*internal variable*)
	END_VAR
END_FUNCTION_BLOCK

FUNCTION_BLOCK MC_BR_InitReceiveNetworkData (*initializes receiving of 4-Byte data from a network station*)
	VAR_INPUT
		Axis : UDINT; (*axis reference*)
		Execute : BOOL; (*initialize receiving of data at the rising edge*)
		NodeNumber : USINT; (*node number of sending network station*)
		BitOffset : UINT; (*bit offset of the data inside the telegram*)
		DataType : UINT; (*data type of the received data*)
		InterpolationMode : USINT; (*interpolation mode of value on receiving drive*)
		ReceiveChannel : USINT; (*receive channel on which the data should be read*)
	END_VAR
	VAR_OUTPUT
		Done : BOOL; (*receiving of data initialized*)
		Busy : BOOL; (*function block is not finished*)
		Error : BOOL; (*error occurred in FB*)
		ErrorID : UINT; (*error number*)
		ReceiveParID : UINT; (*ParID on drive that holds received value*)
	END_VAR
	VAR
		C_Axis : UDINT; (*internal variable*)
		IS : MC_0115_IS_TYP; (*internal variable*)
	END_VAR
END_FUNCTION_BLOCK

FUNCTION_BLOCK MC_BR_InitReceiveNetworkEnc (*initializes receiving of an encoder over the network*)
	VAR_INPUT
		Axis : UDINT; (*axis reference*)
		Execute : BOOL; (*initialize receiving of data at the rising edge*)
		EncoderInformation : MC_NET_ENC_INFO_REF; (*information about the encoder*)
		EncoderParameters : MC_NET_ENC_PARAM_REF; (*parameters for the encoder*)
        ReceiveConfiguration : MC_NET_ENC_CONFIG_REF; (*configuration for processing received encoder values*)
	END_VAR
	VAR_OUTPUT
		Done : BOOL; (*receiving of data initialized*)
		Busy : BOOL; (*function block is not finished*)
		Error : BOOL; (*error occurred in FB*)
		ErrorID : UINT; (*error number*)
		PositionParID : UINT; (*ParID on drive that holds evaluated encoder position*)
	END_VAR
	VAR
		C_Axis : UDINT; (*internal variable*)
		IS : MC_0141_IS_TYP; (*internal variable*)
	END_VAR
END_FUNCTION_BLOCK

FUNCTION_BLOCK MC_BR_InitReceiveParID (*initializes receiving of a ParID on a drive*)
	VAR_INPUT
		Master : UDINT; (*axis reference*)
		Slave : UDINT; (*axis reference*)
		Execute : BOOL; (*initialize receiving of ParID at the rising edge*)
		ParID : UINT; (*ParID that should be received by the drive*)
		InterpolationMode : USINT; (*interpolation mode of value on receiving drive*)
		SendChannel : USINT; (*send channel on which the ParID is sent*)
		ReceiveChannel : USINT; (*receive channel on which the ParID should be read*)
	END_VAR
	VAR_OUTPUT
		Done : BOOL; (*receiving of ParID initialized*)
		Busy : BOOL; (*function block is not finished*)
		Error : BOOL; (*error occurred in FB*)
		ErrorID : UINT; (*error number*)
		ReceiveParID : UINT; (*ParID on slave axis drive that holds received value*)
	END_VAR
	VAR
		C_Master : UDINT; (*internal variable*)
		C_Slave : UDINT; (*internal variable*)
		IS : MC_0112_IS_TYP; (*internal variable*)
	END_VAR
END_FUNCTION_BLOCK

FUNCTION_BLOCK MC_BR_InitSendParID (*initializes sending of a ParID on a drive*)
	VAR_INPUT
		Axis : UDINT; (*axis reference*)
		Execute : BOOL; (*initialize sending of ParID at the rising edge*)
		ParID : UINT; (*ParID that should be sent by the drive*)
		SendChannel : USINT; (*send channel on which the ParID should be sent*)
	END_VAR
	VAR_OUTPUT
		Done : BOOL; (*sending of ParID initialized*)
		Busy : BOOL; (*function block is not finished*)
		Error : BOOL; (*error occurred in FB*)
		ErrorID : UINT; (*error number*)
		AssignedSendChannel : USINT; (*automatically assigned send channel*)
	END_VAR
	VAR
		C_Axis : UDINT; (*internal variable*)
		IS : MC_0111_IS_TYP; (*internal variable*)
	END_VAR
END_FUNCTION_BLOCK

FUNCTION_BLOCK MC_BR_JogVelocity (*enables and executes jog movements*)
	VAR_INPUT
		Axis : UDINT; (*axis reference*)
		Enable : BOOL; (*enables execution of jog movements*)
		Velocity : REAL; (*maximum velocity*)
		Acceleration : REAL; (*maximum acceleration*)
		Deceleration : REAL; (*maximum deceleration*)
		JogPositive : BOOL; (*executes positive movement at high level*)
		JogNegative : BOOL; (*executes negative movement at high level*)
	END_VAR
	VAR_OUTPUT
		Active : BOOL; (*function block is active*)
		Busy : BOOL; (*function block is not finished*)
		CommandAborted : BOOL; (*function block is aborted by another command*)
		Error : BOOL; (*error occurred in FB*)
		ErrorID : UINT; (*error number*)
		Jogging : BOOL; (*jog movement is active*)
	END_VAR
	VAR
		C_Axis : UDINT; (*internal variable*)
		IS : MC_0118_IS_TYP; (*internal variable*)
	END_VAR
END_FUNCTION_BLOCK

FUNCTION_BLOCK MC_BR_JogLimitPosition (*enables and executes jog movements between two limit positions*)
	VAR_INPUT
		Axis : UDINT; (*axis reference*)
		Enable : BOOL; (*enables execution of jog movements*)
		Velocity : REAL; (*maximum velocity*)
		Acceleration : REAL; (*maximum acceleration*)
		Deceleration : REAL; (*maximum deceleration*)
		FirstPosition : REAL; (*lower limit position*)
		LastPosition : REAL; (*higher limit position*)
		JogPositive : BOOL; (*executes positive movement at high level*)
		JogNegative : BOOL; (*executes negative movement at high level*)
	END_VAR
	VAR_OUTPUT
		Active : BOOL; (*function block is active*)
		Busy : BOOL; (*function block is not finished*)
		CommandAborted : BOOL; (*function block is aborted by another command*)
		Error : BOOL; (*error occurred in FB*)
		ErrorID : UINT; (*error number*)
		Jogging : BOOL; (*jog movement is active*)
		LimitReached : BOOL; (*limit position is reached*)
	END_VAR
	VAR
		C_Axis : UDINT; (*internal variable*)
		IS : MC_0119_IS_TYP; (*internal variable*)
	END_VAR
END_FUNCTION_BLOCK

FUNCTION_BLOCK MC_BR_JogTargetPosition (*enables and executes jog movements with a defined target position*)
	VAR_INPUT
		Axis : UDINT; (*axis reference*)
		Enable : BOOL; (*enables executeion of jog movements*)
		Velocity : REAL; (*maximum velocity*)
		Acceleration : REAL; (*maximum acceleration*)
		Deceleration : REAL; (*maximum deceleration*)
		TargetPosition : REAL; (*target position*)
		JogToTarget : BOOL; (*moves to target position at high level*)
		JogPositive : BOOL; (*executes positive movement at high level*)
		JogNegative : BOOL; (*executes negative movement at high level*)
	END_VAR
	VAR_OUTPUT
		Active : BOOL; (*function block is active*)
		Busy : BOOL; (*function block is not finished*)
		CommandAborted : BOOL; (*function block is aborted by another command*)
		Error : BOOL; (*error occurred in FB*)
		ErrorID : UINT; (*error number*)
		Jogging : BOOL; (*jog movement is acitve*)
		MovingToTarget : BOOL; (*axis is moveing to target*)
		TargetReached : BOOL; (*target is reached*)
	END_VAR
	VAR
		C_Axis : UDINT; (*internal variable*)
		IS : MC_0120_IS_TYP; (*internal variable*)
	END_VAR
END_FUNCTION_BLOCK

FUNCTION_BLOCK MC_BR_LimitLoad (*limits the motor torque to set values*)
	VAR_INPUT
		Axis : UDINT; (*axis reference*)
		Enable : BOOL; (*when set limitation is activated*)
		InitData : BOOL; (*initialize the input data*)
		LoadPosAccel : REAL; (*limit value for the motor torque [Nm]*)
		LoadPosDecel : REAL; (*limit value for the motor torque [Nm]*)
		LoadNegAccel : REAL; (*limit value for the motor torque [Nm]*)
		LoadNegDecel : REAL; (*limit value for the motor torque [Nm]*)
		Mode : USINT; (*mode for torque limitation*)
		AdvancedParameters : MC_ADV_LIMITLOAD_REF; (*advanced parameters for torque limitation*)
	END_VAR
	VAR_OUTPUT
		Busy : BOOL; (*function block is not finished*)
		Ready : BOOL; (*parameters initialized*)
		Active : BOOL; (*torque is limited*)
		Error : BOOL; (*error occurred in FB*)
		ErrorID : UINT; (*error number*)
		DataInitialized : BOOL; (*input data initialized*)
	END_VAR
	VAR
		C_Axis : UDINT; (*internal variable*)
		IS : MC_0134_IS_TYP; (*internal variable*)
	END_VAR
END_FUNCTION_BLOCK

FUNCTION_BLOCK MC_BR_LimitLoadCam (*limits the motor torque to value from cam profile*)
	VAR_INPUT
		Axis : UDINT; (*axis reference*)
		Enable : BOOL; (*when set limitation is activated*)
		InitData : BOOL; (*initialize the input data*)
		CamProfileIndexPos : UINT; (*index of cam profile for positive direction*)
		PositionFactorPos : DINT; (*position multiplication factor of cam profile for positive direction*)
		LoadFactorPos : DINT; (*load multiplication factor of cam profile for positive direction*)
		CamProfileIndexNeg : UINT; (*index of cam profile for negative direction*)
		PositionFactorNeg : DINT; (*position multiplication factor of cam profile for negative direction*)
		LoadFactorNeg : DINT; (*load multiplication factor of cam profile for negative direction*)
		Mode : USINT; (*mode for torque limitation*)
	END_VAR
	VAR_OUTPUT
		Busy : BOOL; (*function block is not finished*)
		Ready : BOOL; (*parameters initialized*)
		Active : BOOL; (*torque is limited*)
		Error : BOOL; (*error occurred in FB*)
		ErrorID : UINT; (*error number*)
		DataInitialized : BOOL; (*input data initialized*)
	END_VAR
	VAR
		C_Axis : UDINT; (*internal variable*)
		IS : MC_0135_IS_TYP; (*internal variable*)
	END_VAR
END_FUNCTION_BLOCK

FUNCTION_BLOCK MC_BR_LoadAxisPar (*loads axis parameter from a specified init parameter module to the axis data structure*)
	VAR_INPUT
		Axis : UDINT; (*axis reference*)
		Execute : BOOL; (*loads the init parameter module at rising edge*)
		DataObjectName : STRING[12]; (*name of the init parameter module*)
	END_VAR
	VAR_OUTPUT
		Done : BOOL; (*loading the data is finished*)
		Busy : BOOL; (*function block is not finished*)
		Error : BOOL; (*error occurred in FB*)
		ErrorID : UINT; (*error number*)
	END_VAR
	VAR
		C_Axis : UDINT; (*internal variable*)
		C_DataObjectName : STRING[12]; (*internal variable*)
		state : USINT; (*internal variable*)
		LockIDPar : USINT; (*internal variable*)
		C_ErrorID : UINT; (*internal variable*)
		C_Error : BOOL; (*internal variable*)
		pInit : REFERENCE TO USINT; (*internal variable*)
		pError : REFERENCE TO USINT; (*internal variable*)
	END_VAR
END_FUNCTION_BLOCK

FUNCTION_BLOCK MC_BR_MoveAbsoluteTriggStop (*starts a movement to specified Position, at trigger event it moves the TriggerDistance*)
	VAR_INPUT
		Axis : UDINT; (*axis reference*)
		Execute : BOOL; (*start movement at rising edge*)
		TriggerInput : MC_TRIGGER_REF; (*trigger input signal source*)
		Position : REAL; (*target position for the motion*)
		Velocity : REAL; (*maximum velocity*)
		Acceleration : REAL; (*maximum acceleration*)
		Deceleration : REAL; (*maximum deceleration*)
		Direction : USINT; (*movement direction*)
		TriggerDistance : REAL; (*distance after trigger signal*)
		ForceTriggerDistance : BOOL; (*move trigger distance, even when target position is exceeded*)
	END_VAR
	VAR_OUTPUT
		Done : BOOL; (*absolute move stopped after trigger event or commanded position reached*)
		Busy : BOOL; (*function block is not finished*)
		CommandAborted : BOOL; (*function block is aborted by another command*)
		Error : BOOL; (*error occurred in FB*)
		ErrorID : UINT; (*error number*)
	END_VAR
	VAR
		C_Axis : UDINT; (*internal variable*)
		C_Position : DINT; (*internal variable*)
		C_Velocity : REAL; (*internal variable*)
		C_Acceleration : REAL; (*internal variable*)
		C_Deceleration : REAL; (*internal variable*)
		C_TriggerDistance : DINT; (*internal variable*)
		C_TriggerInput : MC_TRIGGER_REF; (*internal variable*)
		C_ForceTriggerDistance : BOOL; (*internal variable*)
		C_Execute : BOOL; (*internal variable*)
		cmdExecute : BOOL; (*internal variable*)
		C_Direction : USINT; (*internal variable*)
		C_Done : BOOL; (*internal variable*)
		C_CommandAborted : BOOL; (*internal variable*)
		C_Error : BOOL; (*internal variable*)
		C_ErrorID : UINT; (*internal variable*)
		C_CommandedOffset : DINT; (*internal variable*)
		state : USINT; (*internal variable*)
		LockIDPar : USINT; (*internal variable*)
		MoveID : USINT; (*internal variable*)
		oldMoveID : USINT; (*internal variable*)
	END_VAR
END_FUNCTION_BLOCK

FUNCTION_BLOCK MC_BR_MoveAdditiveTriggStop (*starts a movement for the specified distance, at trigger event it moves the TriggerDistance*)
	VAR_INPUT
		Axis : UDINT; (*axis reference*)
		Execute : BOOL; (*start movement at rising edge*)
		TriggerInput : MC_TRIGGER_REF; (*trigger input signal source*)
		Distance : REAL; (*relative distance for the motion*)
		Velocity : REAL; (*value of maximum velocity*)
		Acceleration : REAL; (*value of maximum acceleration*)
		Deceleration : REAL; (*value of maximum deceleration*)
		TriggerDistance : REAL; (*distance after trigger signal*)
		ForceTriggerDistance : BOOL; (*move trigger distance, even when target position is exceeded*)
	END_VAR
	VAR_OUTPUT
		Done : BOOL; (*absolute move stopped after trigger event or commanded position reached*)
		Busy : BOOL; (*function block not finished*)
		CommandAborted : BOOL; (*function block aborted by another command*)
		Error : BOOL; (*error occurred in FB*)
		ErrorID : UINT; (*error number*)
	END_VAR
	VAR
		C_Axis : UDINT; (*internal variable*)
		C_Distance : DINT; (*internal variable*)
		C_Velocity : REAL; (*internal variable*)
		C_Acceleration : REAL; (*internal variable*)
		C_Deceleration : REAL; (*internal variable*)
		C_TriggerDistance : DINT; (*internal variable*)
		C_TriggerInput : MC_TRIGGER_REF; (*internal variable*)
		C_ForceTriggerDistance : BOOL; (*internal variable*)
		C_Execute : BOOL; (*internal variable*)
		cmdExecute : BOOL; (*internal variable*)
		C_Done : BOOL; (*internal variable*)
		C_CommandAborted : BOOL; (*internal variable*)
		C_ErrorID : UINT; (*internal variable*)
		C_Error : BOOL; (*internal variable*)
		state : USINT; (*internal variable*)
		C_CommandedOffset : DINT; (*internal variable*)
		C_CommandedPosition : REAL; (*internal variable*)
		LockIDPar : USINT; (*internal variable*)
		MoveID : USINT; (*internal variable*)
		oldMoveID : USINT; (*internal variable*)
		reserve : USINT; (*internal variable*)
	END_VAR
END_FUNCTION_BLOCK

FUNCTION_BLOCK MC_BR_MoveCyclicPosition (*commands the axis to follow a cyclically transferred position*)
	VAR_INPUT
		Axis : UDINT; (*axis reference*)
		Enable : BOOL; (*as long as Enable is TRUE the cyclic position is transferred to the axis*)
		CyclicPosition : MC_CYCLIC_POSITION; (*cyclic position that is transferred to the axis*)
		Velocity : REAL; (*value of maximum velocity to reach the position*)
		Acceleration : REAL; (*value of maximum acceleration to reach the position*)
		Deceleration : REAL; (*value of maximum deceleration to reach the position*)
		PositionParID : UINT; (*use this ParID as position source instead of CyclicPosition input*)
	END_VAR
	VAR_OUTPUT
		Valid : BOOL; (*position is beeing transferred to the axis*)
		Busy : BOOL; (*function block is not finished*)
		CommandAborted : BOOL; (*function block is aborted by another command*)
		Error : BOOL; (*error occurred in FB*)
		ErrorID : UINT; (*error number*)
		ReceiveParID : UINT; (*ParID that receives the cyclic position*)
	END_VAR
	VAR
		C_Axis : UDINT; (*internal variable*)
		Reserve : USINT; (*internal variable*)
		IS : MC_0081_IS_TYP; (*internal variable*)
	END_VAR
END_FUNCTION_BLOCK

FUNCTION_BLOCK MC_BR_MoveCyclicPositionExt (*commands the axis to follow a cyclically transferred position*)
	VAR_INPUT
		Axis : UDINT; (*axis reference*)
		Enable : BOOL; (*as long as Enable is TRUE the cyclic position is transferred to the axis*)
		CyclicPosition : MC_CYCLIC_POSITION_REF; (*cyclic position that is transferred to the axis*)
		InterpolationMode : USINT; (*interpolation mode of cyclic position on receiving drive*)
		AdvancedParameters : MC_ADVANCED_MOVE_CYC_REF; (*structure for using additional functions*)
	END_VAR
	VAR_OUTPUT
		Valid : BOOL; (*position is beeing transferred to the axis*)
		Busy : BOOL; (*function block is not finished*)
		CommandAborted : BOOL; (*function block is aborted by another command*)
		Error : BOOL; (*error occurred in FB*)
		ErrorID : UINT; (*error number*)
		ReceiveParID : UINT; (*ParID that receives the cyclic position*)
	END_VAR
	VAR
		C_Axis : UDINT; (*internal variable*)
		IS : MC_0124_IS_TYP; (*internal variable*)
	END_VAR
END_FUNCTION_BLOCK

FUNCTION_BLOCK MC_BR_MoveCyclicVelocity (*commands the axis to move with a cyclically transferred velocity*)
	VAR_INPUT
		Axis : UDINT; (*axis reference*)
		Enable : BOOL; (*as long as Enable is TRUE the cyclic velocity is transferred to the axis*)
		CyclicVelocity : REAL; (*cyclic velocity that is transferred to the axis*)
		Direction : USINT; (*direction of movement*)
		Acceleration : REAL; (*value of maximum acceleration to reach the velocity*)
		Deceleration : REAL; (*value of maximum deceleration to reach the velocity*)
		VelocityParID : UINT; (*use this ParID as velocity source instead of CyclicVelocity input*)
	END_VAR
	VAR_OUTPUT
		Valid : BOOL; (*velocity is beeing transferred to the axis*)
		Busy : BOOL; (*function block is not finished*)
		CommandAborted : BOOL; (*function block is aborted by another command*)
		Error : BOOL; (*error occurred in function block*)
		ErrorID : UINT; (*error number*)
		ReceiveParID : UINT; (*ParId that receives the cyclic velocity*)
	END_VAR
	VAR
		C_Axis : UDINT; (*internal variable*)
		IS : MC_0092_IS_TYP; (*internal variable*)
	END_VAR
END_FUNCTION_BLOCK

FUNCTION_BLOCK MC_BR_MoveCyclicVelocityExt (*commands the axis to move with a cyclically transferred velocity*)
	VAR_INPUT
		Axis : UDINT; (*axis reference*)
		Enable : BOOL; (*as long as Enable is TRUE the cyclic velocity is transferred to the axis*)
		CyclicVelocity : REAL; (*cyclic velocity that is transferred to the axis*)
		Direction : USINT; (*direction of movement*)
		InterpolationMode : USINT; (*interpolation mode of cyclic position on receiving drive*)
		AdvancedParameters : MC_ADVANCED_MOVE_CYC_REF; (*structure for using additional functions*)
	END_VAR
	VAR_OUTPUT
		Valid : BOOL; (*velocity is beeing transferred to the axis*)
		Busy : BOOL; (*function block is not finished*)
		CommandAborted : BOOL; (*function block is aborted by another command*)
		Error : BOOL; (*error occurred in function block*)
		ErrorID : UINT; (*error number*)
		ReceiveParID : UINT; (*ParId that receives the cyclic velocity*)
	END_VAR
	VAR
		C_Axis : UDINT; (*internal variable*)
		IS : MC_0125_IS_TYP; (*internal variable*)
	END_VAR
END_FUNCTION_BLOCK

FUNCTION_BLOCK MC_BR_MoveVelocityTriggStop (*starts a movement with specified velocity in specified direction, a trigger stops the axis*)
	VAR_INPUT
		Axis : UDINT; (*axis reference*)
		Execute : BOOL; (*start movement at rising edge*)
		TriggerInput : MC_TRIGGER_REF; (*trigger input signal source*)
		Velocity : REAL; (*maximum velocity*)
		Acceleration : REAL; (*maximum acceleration*)
		Deceleration : REAL; (*maximum deceleration*)
		Direction : USINT; (*movement direction*)
		TriggerDistance : REAL; (*distance after trigger event*)
	END_VAR
	VAR_OUTPUT
		Done : BOOL; (*velocity move stopped after trigger event*)
		Busy : BOOL; (*function block is not finished*)
		CommandAborted : BOOL; (*function block aborted by another command*)
		Error : BOOL; (*error occurred in FB*)
		ErrorID : UINT; (*error number*)
	END_VAR
	VAR
		C_Axis : UDINT; (*internal variable*)
		C_Velocity : REAL; (*internal variable*)
		C_Acceleration : REAL; (*internal variable*)
		C_Deceleration : REAL; (*internal variable*)
		C_Execute : BOOL; (*internal variable*)
		cmdExecute : BOOL; (*internal variable*)
		C_Direction : USINT; (*internal variable*)
		C_Done : BOOL; (*internal variable*)
		C_ErrorID : UINT; (*internal variable*)
		C_CommandAborted : BOOL; (*internal variable*)
		C_Error : BOOL; (*internal variable*)
		C_TriggerInput : MC_TRIGGER_REF; (*internal variable*)
		state : USINT; (*internal variable*)
		C_TriggerDistance : DINT; (*internal variable*)
		LockIDPar : USINT; (*internal variable*)
		MoveID : USINT; (*internal variable*)
		oldMoveID : USINT; (*internal variable*)
		reserve : USINT; (*internal variable*)
	END_VAR
END_FUNCTION_BLOCK

FUNCTION_BLOCK MC_BR_NetTrace (*controls the network command trace*)
	VAR_INPUT
		Execute : BOOL; (*execute command at rising edge*)
		Command : UINT; (*select the command for the network command trace*)
		Configuration : MC_NETTRACECONFIG_REF; (*FB configuration*)
	END_VAR
	VAR_OUTPUT
		Done : BOOL; (*command executed*)
		Busy : BOOL; (*function block is not finished*)
		Error : BOOL; (*error occurred in FB*)
		ErrorID : UINT; (*error number*)
		ErrorRecord : MC_ERRORRECORD_REF; (*error messages that can occur after executing the command*)
	END_VAR
	VAR
		IS : MC_0078_IS_TYP; (*internal variable*)
	END_VAR
END_FUNCTION_BLOCK

FUNCTION_BLOCK MC_BR_NetworkInit (*controls the network initilization*)
	VAR_INPUT
	    Axis : UDINT; (*axis reference*)
		Execute : BOOL; (*execute command at rising edge*)
		Command : UINT; (*select the command for the network initialization*)
	END_VAR
	VAR_OUTPUT
		Done : BOOL; (*command executed*)
		Busy : BOOL; (*function block is not finished*)
		Error : BOOL; (*error occurred in FB*)
		ErrorID : UINT; (*error number*)
	END_VAR
	VAR
		C_Object : UDINT; (*internal variable*)
		IS : MC_0139_IS_TYP; (*internal variable*)
	END_VAR
END_FUNCTION_BLOCK

FUNCTION_BLOCK MC_BR_Offset (*adds an offset to the position of the slave axis*)
	VAR_INPUT
		Slave : UDINT; (*axis reference of the slave axis*)
		Enable : BOOL; (*enable the function block*)
		InitData : BOOL; (*initialize the input data*)
		PerformVelocityControl : BOOL; (*enable the phase shift*)
		Shift : REAL; (*offset shift value*)
		Velocity : REAL; (*velocity for reaching the offset shift*)
		Acceleration : REAL; (*acceleration for reaching the offset shift*)
		ApplicationDistance : REAL; (*distance within which the offset shift occurs*)
		ApplicationMode : UINT; (*basis of movement profile*)
		ShiftMode : UINT; (*definition of how the value on the "Shift" input should be used*)
		AdvancedParameters : MC_ADVANCEDSHIFTPAR_REF; (*structure for using additional functions*)
	END_VAR
	VAR_OUTPUT
		Active : BOOL; (*a offset shift can be executed*)
		Busy : BOOL; (*function block is not finished*)
		Error : BOOL; (*error occurred in FB*)
		ErrorID : UINT; (*error number*)
		ShiftAttained : BOOL; (*offset shift executed*)
		DataInitialized : BOOL; (*input data initialized*)
		ActualShiftValue : REAL; (*current value of shift on the drive*)
	END_VAR
	VAR
		C_Slave : UDINT; (*internal variable*)
		C_InitData : BOOL; (*internal variable*)
		C_PerformVelocityControl : BOOL; (*internal variable*)
		C_Shift : DINT; (*internal variable*)
		C_Velocity : REAL; (*internal variable*)
		C_Acceleration : REAL; (*internal variable*)
		C_ApplicationDistance : DINT; (*internal variable*)
		C_ApplicationMode : UINT; (*internal variable*)
		C_SelectedMaster : UINT; (*internal variable*)
		C_ShiftMode : UINT; (*internal variable*)
		C_AdvancedParameters : MC_ADVANCEDSHIFTPAR_REF; (*internal variable*)
		C_Active : BOOL; (*internal variable*)
		C_Busy : BOOL; (*internal variable*)
		C_Error : BOOL; (*internal variable*)
		C_ErrorID : UINT; (*internal variable*)
		CC_ErrorID : UINT; (*internal variable*)
		C_ShiftAttained : BOOL; (*internal variable*)
		C_DataInitialized : BOOL; (*internal variable*)
		C_AxisState : UINT; (*internal variable*)
		NextState : USINT; (*internal variable*)
		state : USINT; (*internal variable*)
		LockID : USINT; (*internal variable*)
		LockIDPar : USINT; (*internal variable*)
		Factor : UDINT; (*internal variable*)
		RtN : REAL; (*internal variable*)
		VarIndex : UINT; (*internal variable*)
		MpgenIndex : UINT; (*internal variable*)
		C_MpgenStatus : USINT; (*internal variable*)
		MpgenStatusOffset : UINT; (*internal variable*)
		MpgenStatusRecIndex : USINT; (*internal variable*)
		Reserve : USINT; (*internal variable*)
		MpgenValueOffset : UINT; (*internal variable*)
		MpgenValueRecIndex : USINT; (*internal variable*)
		FbID : USINT; (*internal variable*)
		InitDataActive : BOOL; (*internal variable*)
	END_VAR
END_FUNCTION_BLOCK
